Universal Robots URScript: FaiChun_9 Jan_2.script

def Machining2():
  # Default parameters:
  global speed_ms = 0.03
  global speed_rads = 0.75
  global accel_mss = 3
  global accel_radss = 1.2
  global blend_radius_m = 0.0003

  # Add subprograms here
  # Start of main program
  # Program generated by RoboDK v5.6.8 for UR10e on 09/01/2025 15:52:28
  # Using nominal kinematics.
  blend_radius_m = 0.0003
  speed_ms = 0.03
  # set_reference(p[0.335000, -0.075000, 0.000000, 0.000000, 0.000000, 0.000000])
  set_tcp(p[0.000000, 0.000000, 0.252000, 0.000000, 0.000000, 0.000000])
  # Show Tool
  movej([0.564339, -1.115693, -2.614907, -0.981789, 1.570796, 2.135135],accel_radss,speed_rads,0,blend_radius_m)
  movel([0.564339, -1.175740, -2.653333, -0.883316, 1.570796, 2.135135],accel_mss,speed_ms,0,blend_radius_m)
  #SetTool1
  #M_RunCode6
  #SetRPM60000
  speed_ms = 0.01
  #M_RunCode3
  movel([0.564339, -1.203294, -2.667921, -0.841174, 1.570796, 2.135135],accel_mss,speed_ms,0,blend_radius_m)
  speed_ms = 0.003
  movel([0.564339, -1.210543, -2.671504, -0.830343, 1.570796, 2.135135],accel_mss,speed_ms,0,blend_radius_m)
  speed_ms = 0.007
  movel([0.589071, -1.299862, -2.623221, -0.789306, 1.570796, 2.159867],accel_mss,speed_ms,0,blend_radius_m)
  movel([0.580877, -1.304600, -2.620384, -0.787405, 1.570796, 2.151673],accel_mss,speed_ms,0,blend_radius_m)
  movel([0.582153, -1.309303, -2.617539, -0.785547, 1.570796, 2.152950],accel_mss,speed_ms,0,blend_radius_m)
  movel([0.584262, -1.308090, -2.618275, -0.786023, 1.570796, 2.155058],accel_mss,speed_ms,0,blend_radius_m)
  movel([0.583431, -1.304986, -2.620151, -0.787251, 1.570796, 2.154228],accel_mss,speed_ms,0,blend_radius_m)
  movel([0.589492, -1.301500, -2.622244, -0.788646, 1.570796, 2.160288],accel_mss,speed_ms,0,blend_radius_m)
  movel([0.589686, -1.302254, -2.621792, -0.788342, 1.570796, 2.160482],accel_mss,speed_ms,0,blend_radius_m)
  movel([0.590691, -1.306131, -2.619461, -0.786797, 1.570796, 2.161487],accel_mss,speed_ms,0,blend_radius_m)
  movel([0.586616, -1.308460, -2.618051, -0.785878, 1.570796, 2.157412],accel_mss,speed_ms,0,blend_radius_m)
  movel([0.587040, -1.310068, -2.617073, -0.785248, 1.570796, 2.157837],accel_mss,speed_ms,0,blend_radius_m)
  movel([0.591108, -1.307752, -2.618481, -0.786157, 1.570796, 2.161905],accel_mss,speed_ms,0,blend_radius_m)
  movel([0.592288, -1.312350, -2.615680, -0.784359, 1.570796, 2.163085],accel_mss,speed_ms,0,blend_radius_m)
  movel([0.588242, -1.314642, -2.614274, -0.783473, 1.570796, 2.159038],accel_mss,speed_ms,0,blend_radius_m)
  movel([0.589043, -1.317715, -2.612378, -0.782297, 1.570796, 2.159840],accel_mss,speed_ms,0,blend_radius_m)
  movel([0.583100, -1.321078, -2.610288, -0.781023, 1.570796, 2.153897],accel_mss,speed_ms,0,blend_radius_m)
  movel([0.582276, -1.318031, -2.612181, -0.782176, 1.570796, 2.153073],accel_mss,speed_ms,0,blend_radius_m)
  movel([0.580193, -1.319220, -2.611444, -0.781725, 1.570796, 2.150989],accel_mss,speed_ms,0,blend_radius_m)
  movel([0.581023, -1.322259, -2.609550, -0.780580, 1.570796, 2.151819],accel_mss,speed_ms,0,blend_radius_m)
  movel([0.576077, -1.325076, -2.607784, -0.779529, 1.570796, 2.146874],accel_mss,speed_ms,0,blend_radius_m)
  movel([0.575122, -1.325624, -2.607439, -0.779326, 1.570796, 2.145918],accel_mss,speed_ms,0,blend_radius_m)
  movel([0.573856, -1.321163, -2.610235, -0.780991, 1.570796, 2.144653],accel_mss,speed_ms,0,blend_radius_m)
  movel([0.577859, -1.318861, -2.611667, -0.781861, 1.570796, 2.148656],accel_mss,speed_ms,0,blend_radius_m)
  movel([0.577420, -1.317283, -2.612645, -0.782461, 1.570796, 2.148217],accel_mss,speed_ms,0,blend_radius_m)
  movel([0.571335, -1.320792, -2.610466, -0.781131, 1.570796, 2.142131],accel_mss,speed_ms,0,blend_radius_m)
  movel([0.573058, -1.326803, -2.606696, -0.778890, 1.570796, 2.143854],accel_mss,speed_ms,0,blend_radius_m)
  movel([0.470799, -1.388192, -2.565343, -0.758854, 1.570796, 2.041595],accel_mss,speed_ms,0,blend_radius_m)
  movel([0.378716, -1.448552, -2.519372, -0.744466, 1.570796, 1.949513],accel_mss,speed_ms,0,blend_radius_m)
  movel([0.375919, -1.444184, -2.522882, -0.745323, 1.570796, 1.946716],accel_mss,speed_ms,0,blend_radius_m)
  movel([0.371026, -1.447561, -2.520170, -0.744657, 1.570796, 1.941822],accel_mss,speed_ms,0,blend_radius_m)
  movel([0.371758, -1.448686, -2.519263, -0.744440, 1.570796, 1.942554],accel_mss,speed_ms,0,blend_radius_m)
  movel([0.374972, -1.446470, -2.521049, -0.744871, 1.570796, 1.945769],accel_mss,speed_ms,0,blend_radius_m)
  movel([0.377041, -1.449694, -2.518449, -0.744246, 1.570796, 1.947837],accel_mss,speed_ms,0,blend_radius_m)
  movel([0.376268, -1.450223, -2.518020, -0.744145, 1.570796, 1.947064],accel_mss,speed_ms,0,blend_radius_m)
  movel([0.372297, -1.452950, -2.515807, -0.743632, 1.570796, 1.943093],accel_mss,speed_ms,0,blend_radius_m)
  movel([0.370895, -1.450790, -2.517562, -0.744037, 1.570796, 1.941691],accel_mss,speed_ms,0,blend_radius_m)
  movel([0.369236, -1.451936, -2.516632, -0.743821, 1.570796, 1.940032],accel_mss,speed_ms,0,blend_radius_m)
  movel([0.370642, -1.454090, -2.514879, -0.743420, 1.570796, 1.941438],accel_mss,speed_ms,0,blend_radius_m)
  movel([0.365939, -1.457337, -2.512222, -0.742829, 1.570796, 1.936735],accel_mss,speed_ms,0,blend_radius_m)
  movel([0.364521, -1.455203, -2.513970, -0.743216, 1.570796, 1.935317],accel_mss,speed_ms,0,blend_radius_m)
  movel([0.361355, -1.457405, -2.512167, -0.742817, 1.570796, 1.932152],accel_mss,speed_ms,0,blend_radius_m)
  movel([0.359234, -1.454259, -2.514741, -0.743389, 1.570796, 1.930031],accel_mss,speed_ms,0,blend_radius_m)
  movel([0.362410, -1.452037, -2.516550, -0.743802, 1.570796, 1.933206],accel_mss,speed_ms,0,blend_radius_m)
  movel([0.361665, -1.450927, -2.517450, -0.744011, 1.570796, 1.932462],accel_mss,speed_ms,0,blend_radius_m)
  movel([0.358487, -1.453153, -2.515642, -0.743594, 1.570796, 1.929284],accel_mss,speed_ms,0,blend_radius_m)
  movel([0.356688, -1.450515, -2.517784, -0.744090, 1.570796, 1.927484],accel_mss,speed_ms,0,blend_radius_m)
  movel([0.356339, -1.450002, -2.518199, -0.744187, 1.570796, 1.927136],accel_mss,speed_ms,0,blend_radius_m)
  movel([0.361066, -1.446678, -2.520881, -0.744830, 1.570796, 1.931863],accel_mss,speed_ms,0,blend_radius_m)
  movel([0.362508, -1.448824, -2.519152, -0.744413, 1.570796, 1.933304],accel_mss,speed_ms,0,blend_radius_m)
  movel([0.364168, -1.447664, -2.520088, -0.744637, 1.570796, 1.934964],accel_mss,speed_ms,0,blend_radius_m)
  movel([0.361980, -1.444391, -2.522716, -0.745282, 1.570796, 1.932777],accel_mss,speed_ms,0,blend_radius_m)
  movel([0.355583, -1.448897, -2.519093, -0.744399, 1.570796, 1.926379],accel_mss,speed_ms,0,blend_radius_m)
  movel([0.355230, -1.448386, -2.519506, -0.744497, 1.570796, 1.926027],accel_mss,speed_ms,0,blend_radius_m)
  movel([0.312755, -1.390773, -2.563487, -0.758128, 1.570796, 1.883551],accel_mss,speed_ms,0,blend_radius_m)
  movel([0.262445, -1.332364, -2.603164, -0.776861, 1.570796, 1.833241],accel_mss,speed_ms,0,blend_radius_m)
  movel([0.269473, -1.326239, -2.607051, -0.779098, 1.570796, 1.840270],accel_mss,speed_ms,0,blend_radius_m)
  movel([0.266416, -1.322928, -2.609132, -0.780329, 1.570796, 1.837212],accel_mss,speed_ms,0,blend_radius_m)
  movel([0.264580, -1.324533, -2.608125, -0.779731, 1.570796, 1.835377],accel_mss,speed_ms,0,blend_radius_m)
  movel([0.266599, -1.326703, -2.606759, -0.778927, 1.570796, 1.837395],accel_mss,speed_ms,0,blend_radius_m)
  movel([0.261398, -1.331241, -2.603881, -0.777267, 1.570796, 1.832194],accel_mss,speed_ms,0,blend_radius_m)
  movel([0.260914, -1.330724, -2.604210, -0.777455, 1.570796, 1.831710],accel_mss,speed_ms,0,blend_radius_m)
  movel([0.258394, -1.328064, -2.605899, -0.778426, 1.570796, 1.829190],accel_mss,speed_ms,0,blend_radius_m)
  movel([0.261907, -1.324978, -2.607845, -0.779565, 1.570796, 1.832703],accel_mss,speed_ms,0,blend_radius_m)
  movel([0.260849, -1.323857, -2.608550, -0.779982, 1.570796, 1.831646],accel_mss,speed_ms,0,blend_radius_m)
  movel([0.257334, -1.326952, -2.606602, -0.778835, 1.570796, 1.828131],accel_mss,speed_ms,0,blend_radius_m)
  movel([0.254293, -1.323782, -2.608597, -0.780010, 1.570796, 1.825090],accel_mss,speed_ms,0,blend_radius_m)
  movel([0.257815, -1.320661, -2.610547, -0.781180, 1.570796, 1.828612],accel_mss,speed_ms,0,blend_radius_m)
  movel([0.255752, -1.318503, -2.611889, -0.781997, 1.570796, 1.826548],accel_mss,speed_ms,0,blend_radius_m)
  movel([0.261012, -1.313833, -2.614771, -0.783785, 1.570796, 1.831808],accel_mss,speed_ms,0,blend_radius_m)
  movel([0.263069, -1.316016, -2.613428, -0.782946, 1.570796, 1.833865],accel_mss,speed_ms,0,blend_radius_m)
  movel([0.264921, -1.314382, -2.614434, -0.783573, 1.570796, 1.835718],accel_mss,speed_ms,0,blend_radius_m)
  movel([0.262867, -1.312190, -2.615778, -0.784421, 1.570796, 1.833663],accel_mss,speed_ms,0,blend_radius_m)
  movel([0.267321, -1.308250, -2.618179, -0.785961, 1.570796, 1.838117],accel_mss,speed_ms,0,blend_radius_m)
  movel([0.268189, -1.307485, -2.618642, -0.786262, 1.570796, 1.838985],accel_mss,speed_ms,0,blend_radius_m)
  movel([0.271218, -1.310771, -2.616645, -0.784973, 1.570796, 1.842014],accel_mss,speed_ms,0,blend_radius_m)
  movel([0.267627, -1.313924, -2.614715, -0.783750, 1.570796, 1.838423],accel_mss,speed_ms,0,blend_radius_m)
  movel([0.268684, -1.315067, -2.614012, -0.783310, 1.570796, 1.839480],accel_mss,speed_ms,0,blend_radius_m)
  movel([0.274144, -1.310287, -2.616940, -0.785162, 1.570796, 1.844940],accel_mss,speed_ms,0,blend_radius_m)
  movel([0.270069, -1.305826, -2.619645, -0.786918, 1.570796, 1.840865],accel_mss,speed_ms,0,blend_radius_m)
  movel([0.376357, -1.214643, -2.669493, -0.828252, 1.570796, 1.947154],accel_mss,speed_ms,0,blend_radius_m)
  movel([0.499980, -1.114188, -2.713609, -0.884591, 1.570796, 2.070776],accel_mss,speed_ms,0,blend_radius_m)
  movel([0.501179, -1.113243, -2.713976, -0.885169, 1.570796, 2.071975],accel_mss,speed_ms,0,blend_radius_m)
  movel([0.504077, -1.120540, -2.711120, -0.880729, 1.570796, 2.074873],accel_mss,speed_ms,0,blend_radius_m)
  movel([0.511634, -1.114642, -2.713433, -0.884314, 1.570796, 2.082430],accel_mss,speed_ms,0,blend_radius_m)
  movel([0.510904, -1.112724, -2.714178, -0.885487, 1.570796, 2.081700],accel_mss,speed_ms,0,blend_radius_m)
  movel([0.505914, -1.116627, -2.712658, -0.883104, 1.570796, 2.076710],accel_mss,speed_ms,0,blend_radius_m)
  movel([0.503784, -1.111195, -2.714769, -0.886425, 1.570796, 2.074581],accel_mss,speed_ms,0,blend_radius_m)
  movel([0.504986, -1.110247, -2.715135, -0.887007, 1.570796, 2.075782],accel_mss,speed_ms,0,blend_radius_m)
  movel([0.511228, -1.105329, -2.717019, -0.890042, 1.570796, 2.082024],accel_mss,speed_ms,0,blend_radius_m)
  movel([0.512639, -1.109056, -2.715593, -0.887740, 1.570796, 2.083436],accel_mss,speed_ms,0,blend_radius_m)
  movel([0.515254, -1.107012, -2.716376, -0.889001, 1.570796, 2.086050],accel_mss,speed_ms,0,blend_radius_m)
  movel([0.513852, -1.103266, -2.717802, -0.891321, 1.570796, 2.084649],accel_mss,speed_ms,0,blend_radius_m)
  movel([0.521382, -1.097360, -2.720023, -0.895006, 1.570796, 2.092179],accel_mss,speed_ms,0,blend_radius_m)
  movel([0.522759, -1.101158, -2.718598, -0.892633, 1.570796, 2.093556],accel_mss,speed_ms,0,blend_radius_m)
  movel([0.527861, -1.097189, -2.720087, -0.895113, 1.570796, 2.098658],accel_mss,speed_ms,0,blend_radius_m)
  movel([0.529846, -1.102848, -2.717960, -0.891581, 1.570796, 2.100643],accel_mss,speed_ms,0,blend_radius_m)
  movel([0.524769, -1.106765, -2.716471, -0.889153, 1.570796, 2.095565],accel_mss,speed_ms,0,blend_radius_m)
  movel([0.525468, -1.108724, -2.715721, -0.887945, 1.570796, 2.096264],accel_mss,speed_ms,0,blend_radius_m)
  movel([0.530535, -1.104825, -2.717210, -0.890354, 1.570796, 2.101331],accel_mss,speed_ms,0,blend_radius_m)
  movel([0.532478, -1.110454, -2.715055, -0.886880, 1.570796, 2.103274],accel_mss,speed_ms,0,blend_radius_m)
  movel([0.525035, -1.116137, -2.712849, -0.883402, 1.570796, 2.095831],accel_mss,speed_ms,0,blend_radius_m)
  movel([0.523692, -1.112395, -2.714305, -0.885689, 1.570796, 2.094489],accel_mss,speed_ms,0,blend_radius_m)
  movel([0.521088, -1.114399, -2.713527, -0.884462, 1.570796, 2.091884],accel_mss,speed_ms,0,blend_radius_m)
  movel([0.523134, -1.120056, -2.711311, -0.881022, 1.570796, 2.093931],accel_mss,speed_ms,0,blend_radius_m)
  movel([0.533154, -1.112420, -2.714296, -0.885673, 1.570796, 2.103950],accel_mss,speed_ms,0,blend_radius_m)
  movel([0.564339, -1.210543, -2.671504, -0.830343, 1.570796, 2.135135],accel_mss,speed_ms,0,blend_radius_m)
  speed_ms = 0.003
  movel([0.564339, -1.203294, -2.667921, -0.841174, 1.570796, 2.135135],accel_mss,speed_ms,0,blend_radius_m)
  speed_ms = 0.03
  movel([0.564339, -1.175740, -2.653333, -0.883316, 1.570796, 2.135135],accel_mss,speed_ms,0,blend_radius_m)
  #M_RunCode9
  movel([0.508673, -1.124915, -2.675707, -0.911767, 1.570796, 2.079469],accel_mss,speed_ms,0,blend_radius_m)
  #M_RunCode3
  movel([0.508673, -1.152779, -2.690963, -0.868647, 1.570796, 2.079469],accel_mss,speed_ms,0,blend_radius_m)
  speed_ms = 0.003
  movel([0.508673, -1.160141, -2.694716, -0.857531, 1.570796, 2.079469],accel_mss,speed_ms,0,blend_radius_m)
  speed_ms = 0.007
  movel([0.506502, -1.162157, -2.693839, -0.856392, 1.570796, 2.077298],accel_mss,speed_ms,0,blend_radius_m)
  movel([0.504257, -1.163601, -2.693209, -0.855579, 1.570796, 2.075054],accel_mss,speed_ms,0,blend_radius_m)
  movel([0.501934, -1.164482, -2.692823, -0.855084, 1.570796, 2.072730],accel_mss,speed_ms,0,blend_radius_m)
  movel([0.499527, -1.164799, -2.692684, -0.854906, 1.570796, 2.070323],accel_mss,speed_ms,0,blend_radius_m)
  movel([0.497561, -1.164580, -2.692780, -0.855029, 1.570796, 2.068358],accel_mss,speed_ms,0,blend_radius_m)
  movel([0.495980, -1.163844, -2.693102, -0.855442, 1.570796, 2.066776],accel_mss,speed_ms,0,blend_radius_m)
  movel([0.494731, -1.162733, -2.693588, -0.856068, 1.570796, 2.065527],accel_mss,speed_ms,0,blend_radius_m)
  movel([0.493766, -1.161377, -2.694179, -0.856833, 1.570796, 2.064563],accel_mss,speed_ms,0,blend_radius_m)
  movel([0.492038, -1.157449, -2.695881, -0.859059, 1.570796, 2.062834],accel_mss,speed_ms,0,blend_radius_m)
  movel([0.490361, -1.153755, -2.697467, -0.861167, 1.570796, 2.061158],accel_mss,speed_ms,0,blend_radius_m)
  movel([0.489477, -1.152506, -2.698000, -0.861883, 1.570796, 2.060274],accel_mss,speed_ms,0,blend_radius_m)
  movel([0.488348, -1.151492, -2.698432, -0.862465, 1.570796, 2.059144],accel_mss,speed_ms,0,blend_radius_m)
  movel([0.486938, -1.150837, -2.698710, -0.862842, 1.570796, 2.057734],accel_mss,speed_ms,0,blend_radius_m)
  movel([0.485211, -1.150668, -2.698782, -0.862939, 1.570796, 2.056007],accel_mss,speed_ms,0,blend_radius_m)
  movel([0.484699, -1.151781, -2.698309, -0.862299, 1.570796, 2.055495],accel_mss,speed_ms,0,blend_radius_m)
  movel([0.483417, -1.154849, -2.696999, -0.860541, 1.570796, 2.054213],accel_mss,speed_ms,0,blend_radius_m)
  movel([0.482581, -1.157515, -2.695853, -0.859021, 1.570796, 2.053377],accel_mss,speed_ms,0,blend_radius_m)
  movel([0.482187, -1.159786, -2.694871, -0.857732, 1.570796, 2.052983],accel_mss,speed_ms,0,blend_radius_m)
  movel([0.482229, -1.161669, -2.694052, -0.856668, 1.570796, 2.053026],accel_mss,speed_ms,0,blend_radius_m)
  movel([0.482647, -1.163187, -2.693390, -0.855812, 1.570796, 2.053443],accel_mss,speed_ms,0,blend_radius_m)
  movel([0.483386, -1.164368, -2.692873, -0.855148, 1.570796, 2.054183],accel_mss,speed_ms,0,blend_radius_m)
  movel([0.484448, -1.165208, -2.692505, -0.854677, 1.570796, 2.055244],accel_mss,speed_ms,0,blend_radius_m)
  movel([0.485828, -1.165715, -2.692281, -0.854392, 1.570796, 2.056624],accel_mss,speed_ms,0,blend_radius_m)
  movel([0.477331, -1.166016, -2.692149, -0.854224, 1.570796, 2.048127],accel_mss,speed_ms,0,blend_radius_m)
  movel([0.490968, -1.136326, -2.704766, -0.871297, 1.570796, 2.061764],accel_mss,speed_ms,0,blend_radius_m)
  movel([0.491843, -1.136290, -2.704781, -0.871318, 1.570796, 2.062639],accel_mss,speed_ms,0,blend_radius_m)
  movel([0.493898, -1.136547, -2.704675, -0.871167, 1.570796, 2.064694],accel_mss,speed_ms,0,blend_radius_m)
  movel([0.495585, -1.137510, -2.704280, -0.870600, 1.570796, 2.066381],accel_mss,speed_ms,0,blend_radius_m)
  movel([0.496938, -1.138969, -2.703678, -0.869741, 1.570796, 2.067734],accel_mss,speed_ms,0,blend_radius_m)
  movel([0.497990, -1.140717, -2.702955, -0.868716, 1.570796, 2.068786],accel_mss,speed_ms,0,blend_radius_m)
  movel([0.500129, -1.145961, -2.700769, -0.865660, 1.570796, 2.070926],accel_mss,speed_ms,0,blend_radius_m)
  movel([0.502024, -1.150859, -2.698701, -0.862829, 1.570796, 2.072821],accel_mss,speed_ms,0,blend_radius_m)
  movel([0.502966, -1.152496, -2.698005, -0.861888, 1.570796, 2.073762],accel_mss,speed_ms,0,blend_radius_m)
  movel([0.504145, -1.153842, -2.697430, -0.861117, 1.570796, 2.074941],accel_mss,speed_ms,0,blend_radius_m)
  movel([0.505585, -1.154734, -2.697048, -0.860607, 1.570796, 2.076381],accel_mss,speed_ms,0,blend_radius_m)
  movel([0.507301, -1.155017, -2.696927, -0.860445, 1.570796, 2.078097],accel_mss,speed_ms,0,blend_radius_m)
  movel([0.509687, -1.154592, -2.697109, -0.860688, 1.570796, 2.080483],accel_mss,speed_ms,0,blend_radius_m)
  movel([0.510798, -1.154086, -2.697325, -0.860977, 1.570796, 2.081594],accel_mss,speed_ms,0,blend_radius_m)
  movel([0.511860, -1.153380, -2.697627, -0.861382, 1.570796, 2.082656],accel_mss,speed_ms,0,blend_radius_m)
  movel([0.513679, -1.151630, -2.698373, -0.862386, 1.570796, 2.084475],accel_mss,speed_ms,0,blend_radius_m)
  movel([0.514984, -1.149603, -2.699233, -0.863553, 1.570796, 2.085781],accel_mss,speed_ms,0,blend_radius_m)
  movel([0.515524, -1.148232, -2.699813, -0.864344, 1.570796, 2.086320],accel_mss,speed_ms,0,blend_radius_m)
  movel([0.515638, -1.147219, -2.700240, -0.864930, 1.570796, 2.086434],accel_mss,speed_ms,0,blend_radius_m)
  movel([0.515378, -1.146593, -2.700503, -0.865293, 1.570796, 2.086174],accel_mss,speed_ms,0,blend_radius_m)
  movel([0.514794, -1.146390, -2.700588, -0.865411, 1.570796, 2.085591],accel_mss,speed_ms,0,blend_radius_m)
  movel([0.513538, -1.146896, -2.700375, -0.865117, 1.570796, 2.084335],accel_mss,speed_ms,0,blend_radius_m)
  movel([0.512295, -1.147497, -2.700123, -0.864769, 1.570796, 2.083092],accel_mss,speed_ms,0,blend_radius_m)
  movel([0.510910, -1.147730, -2.700025, -0.864635, 1.570796, 2.081706],accel_mss,speed_ms,0,blend_radius_m)
  movel([0.509562, -1.147401, -2.700163, -0.864825, 1.570796, 2.080359],accel_mss,speed_ms,0,blend_radius_m)
  movel([0.508936, -1.146367, -2.700598, -0.865424, 1.570796, 2.079732],accel_mss,speed_ms,0,blend_radius_m)
  movel([0.508971, -1.144842, -2.701238, -0.866310, 1.570796, 2.079767],accel_mss,speed_ms,0,blend_radius_m)
  movel([0.509601, -1.143041, -2.701990, -0.867358, 1.570796, 2.080397],accel_mss,speed_ms,0,blend_radius_m)
  movel([0.510703, -1.141227, -2.702744, -0.868418, 1.570796, 2.081499],accel_mss,speed_ms,0,blend_radius_m)
  movel([0.512151, -1.139669, -2.703389, -0.869331, 1.570796, 2.082947],accel_mss,speed_ms,0,blend_radius_m)
  movel([0.513800, -1.138587, -2.703836, -0.869966, 1.570796, 2.084597],accel_mss,speed_ms,0,blend_radius_m)
  movel([0.515498, -1.138213, -2.703990, -0.870186, 1.570796, 2.086294],accel_mss,speed_ms,0,blend_radius_m)
  movel([0.516742, -1.138401, -2.703913, -0.870075, 1.570796, 2.087539],accel_mss,speed_ms,0,blend_radius_m)
  movel([0.517622, -1.139001, -2.703665, -0.869722, 1.570796, 2.088419],accel_mss,speed_ms,0,blend_radius_m)
  movel([0.518134, -1.140018, -2.703245, -0.869126, 1.570796, 2.088931],accel_mss,speed_ms,0,blend_radius_m)
  movel([0.518284, -1.141439, -2.702656, -0.868294, 1.570796, 2.089081],accel_mss,speed_ms,0,blend_radius_m)
  movel([0.518110, -1.143170, -2.701936, -0.867283, 1.570796, 2.088906],accel_mss,speed_ms,0,blend_radius_m)
  movel([0.517640, -1.145109, -2.701126, -0.866154, 1.570796, 2.088437],accel_mss,speed_ms,0,blend_radius_m)
  movel([0.515835, -1.149598, -2.699236, -0.863556, 1.570796, 2.086632],accel_mss,speed_ms,0,blend_radius_m)
  movel([0.514301, -1.152485, -2.698009, -0.861894, 1.570796, 2.085098],accel_mss,speed_ms,0,blend_radius_m)
  movel([0.512598, -1.155205, -2.696846, -0.860338, 1.570796, 2.083394],accel_mss,speed_ms,0,blend_radius_m)
  movel([0.510722, -1.157753, -2.695750, -0.858886, 1.570796, 2.081518],accel_mss,speed_ms,0,blend_radius_m)
  movel([0.508673, -1.160141, -2.694716, -0.857531, 1.570796, 2.079469],accel_mss,speed_ms,0,blend_radius_m)
  speed_ms = 0.003
  movel([0.508673, -1.152779, -2.690963, -0.868647, 1.570796, 2.079469],accel_mss,speed_ms,0,blend_radius_m)
  speed_ms = 0.03
  movel([0.508673, -1.124915, -2.675707, -0.911767, 1.570796, 2.079469],accel_mss,speed_ms,0,blend_radius_m)
  #M_RunCode9
  movel([0.497081, -1.144256, -2.667496, -0.900636, 1.570796, 2.067877],accel_mss,speed_ms,0,blend_radius_m)
  #M_RunCode3
  movel([0.497081, -1.172027, -2.682500, -0.857862, 1.570796, 2.067877],accel_mss,speed_ms,0,blend_radius_m)
  speed_ms = 0.003
  movel([0.497081, -1.179353, -2.686188, -0.846848, 1.570796, 2.067877],accel_mss,speed_ms,0,blend_radius_m)
  speed_ms = 0.007
  movel([0.498395, -1.179888, -2.685945, -0.846556, 1.570796, 2.069191],accel_mss,speed_ms,0,blend_radius_m)
  movel([0.499154, -1.180637, -2.685604, -0.846148, 1.570796, 2.069950],accel_mss,speed_ms,0,blend_radius_m)
  movel([0.499362, -1.181606, -2.685163, -0.845621, 1.570796, 2.070158],accel_mss,speed_ms,0,blend_radius_m)
  movel([0.499017, -1.182788, -2.684622, -0.844979, 1.570796, 2.069813],accel_mss,speed_ms,0,blend_radius_m)
  movel([0.498226, -1.183973, -2.684079, -0.844337, 1.570796, 2.069022],accel_mss,speed_ms,0,blend_radius_m)
  movel([0.497089, -1.184946, -2.683632, -0.843811, 1.570796, 2.067885],accel_mss,speed_ms,0,blend_radius_m)
  movel([0.495612, -1.185707, -2.683282, -0.843400, 1.570796, 2.066408],accel_mss,speed_ms,0,blend_radius_m)
  movel([0.493784, -1.186265, -2.683025, -0.843099, 1.570796, 2.064581],accel_mss,speed_ms,0,blend_radius_m)
  movel([0.488939, -1.186979, -2.682695, -0.842715, 1.570796, 2.059736],accel_mss,speed_ms,0,blend_radius_m)
  movel([0.482396, -1.187317, -2.682539, -0.842533, 1.570796, 2.053192],accel_mss,speed_ms,0,blend_radius_m)
  movel([0.476031, -1.187267, -2.682562, -0.842560, 1.570796, 2.046827],accel_mss,speed_ms,0,blend_radius_m)
  movel([0.471758, -1.186758, -2.682797, -0.842834, 1.570796, 2.042555],accel_mss,speed_ms,0,blend_radius_m)
  movel([0.470420, -1.186270, -2.683022, -0.843096, 1.570796, 2.041216],accel_mss,speed_ms,0,blend_radius_m)
  movel([0.469629, -1.185561, -2.683349, -0.843479, 1.570796, 2.040426],accel_mss,speed_ms,0,blend_radius_m)
  movel([0.469386, -1.184621, -2.683782, -0.843986, 1.570796, 2.040183],accel_mss,speed_ms,0,blend_radius_m)
  movel([0.469698, -1.183447, -2.684320, -0.844621, 1.570796, 2.040494],accel_mss,speed_ms,0,blend_radius_m)
  movel([0.470461, -1.182257, -2.684865, -0.845267, 1.570796, 2.041257],accel_mss,speed_ms,0,blend_radius_m)
  movel([0.471587, -1.181260, -2.685321, -0.845809, 1.570796, 2.042384],accel_mss,speed_ms,0,blend_radius_m)
  movel([0.473070, -1.180460, -2.685685, -0.846244, 1.570796, 2.043867],accel_mss,speed_ms,0,blend_radius_m)
  movel([0.474917, -1.179854, -2.685960, -0.846575, 1.570796, 2.045714],accel_mss,speed_ms,0,blend_radius_m)
  movel([0.479828, -1.179041, -2.686329, -0.847018, 1.570796, 2.050624],accel_mss,speed_ms,0,blend_radius_m)
  movel([0.486445, -1.178651, -2.686507, -0.847232, 1.570796, 2.057241],accel_mss,speed_ms,0,blend_radius_m)
  movel([0.492832, -1.178747, -2.686463, -0.847179, 1.570796, 2.063629],accel_mss,speed_ms,0,blend_radius_m)
  movel([0.497081, -1.179353, -2.686188, -0.846848, 1.570796, 2.067877],accel_mss,speed_ms,0,blend_radius_m)
  speed_ms = 0.003
  movel([0.497081, -1.172027, -2.682500, -0.857862, 1.570796, 2.067877],accel_mss,speed_ms,0,blend_radius_m)
  speed_ms = 0.03
  movel([0.497081, -1.144256, -2.667496, -0.900636, 1.570796, 2.067877],accel_mss,speed_ms,0,blend_radius_m)
  #M_RunCode9
  movel([0.501396, -1.142283, -2.668351, -0.901755, 1.570796, 2.072192],accel_mss,speed_ms,0,blend_radius_m)
  #M_RunCode3
  movel([0.501396, -1.170065, -2.683380, -0.858944, 1.570796, 2.072192],accel_mss,speed_ms,0,blend_radius_m)
  speed_ms = 0.003
  movel([0.501396, -1.177394, -2.687075, -0.847919, 1.570796, 2.072192],accel_mss,speed_ms,0,blend_radius_m)
  speed_ms = 0.007
  movel([0.501126, -1.179098, -2.686304, -0.846987, 1.570796, 2.071922],accel_mss,speed_ms,0,blend_radius_m)
  movel([0.500589, -1.180897, -2.685486, -0.846006, 1.570796, 2.071385],accel_mss,speed_ms,0,blend_radius_m)
  movel([0.499790, -1.182783, -2.684624, -0.844981, 1.570796, 2.070587],accel_mss,speed_ms,0,blend_radius_m)
  movel([0.498777, -1.184668, -2.683760, -0.843961, 1.570796, 2.069573],accel_mss,speed_ms,0,blend_radius_m)
  movel([0.497593, -1.186454, -2.682938, -0.842998, 1.570796, 2.068389],accel_mss,speed_ms,0,blend_radius_m)
  movel([0.496241, -1.188138, -2.682158, -0.842092, 1.570796, 2.067037],accel_mss,speed_ms,0,blend_radius_m)
  movel([0.494719, -1.189727, -2.681421, -0.841241, 1.570796, 2.065515],accel_mss,speed_ms,0,blend_radius_m)
  movel([0.493045, -1.191188, -2.680740, -0.840460, 1.570796, 2.063841],accel_mss,speed_ms,0,blend_radius_m)
  movel([0.491239, -1.192488, -2.680133, -0.839768, 1.570796, 2.062036],accel_mss,speed_ms,0,blend_radius_m)
  movel([0.489295, -1.193633, -2.679596, -0.839160, 1.570796, 2.060092],accel_mss,speed_ms,0,blend_radius_m)
  movel([0.487213, -1.194624, -2.679131, -0.838635, 1.570796, 2.058010],accel_mss,speed_ms,0,blend_radius_m)
  movel([0.485034, -1.195426, -2.678753, -0.838210, 1.570796, 2.055830],accel_mss,speed_ms,0,blend_radius_m)
  movel([0.482787, -1.196014, -2.678476, -0.837899, 1.570796, 2.053583],accel_mss,speed_ms,0,blend_radius_m)
  movel([0.480475, -1.196388, -2.678299, -0.837702, 1.570796, 2.051271],accel_mss,speed_ms,0,blend_radius_m)
  movel([0.478097, -1.196547, -2.678224, -0.837618, 1.570796, 2.048893],accel_mss,speed_ms,0,blend_radius_m)
  movel([0.475817, -1.196490, -2.678251, -0.837648, 1.570796, 2.046613],accel_mss,speed_ms,0,blend_radius_m)
  movel([0.473808, -1.196212, -2.678382, -0.837795, 1.570796, 2.044604],accel_mss,speed_ms,0,blend_radius_m)
  movel([0.472068, -1.195712, -2.678618, -0.838059, 1.570796, 2.042864],accel_mss,speed_ms,0,blend_radius_m)
  movel([0.470598, -1.194990, -2.678958, -0.838441, 1.570796, 2.041394],accel_mss,speed_ms,0,blend_radius_m)
  movel([0.469404, -1.194073, -2.679390, -0.838926, 1.570796, 2.040200],accel_mss,speed_ms,0,blend_radius_m)
  movel([0.468492, -1.192991, -2.679897, -0.839500, 1.570796, 2.039288],accel_mss,speed_ms,0,blend_radius_m)
  movel([0.467863, -1.191747, -2.680479, -0.840162, 1.570796, 2.038659],accel_mss,speed_ms,0,blend_radius_m)
  movel([0.467519, -1.190332, -2.681140, -0.840918, 1.570796, 2.038316],accel_mss,speed_ms,0,blend_radius_m)
  movel([0.467450, -1.188781, -2.681861, -0.841747, 1.570796, 2.038247],accel_mss,speed_ms,0,blend_radius_m)
  movel([0.467649, -1.187124, -2.682628, -0.842637, 1.570796, 2.038445],accel_mss,speed_ms,0,blend_radius_m)
  movel([0.468121, -1.185356, -2.683444, -0.843589, 1.570796, 2.038917],accel_mss,speed_ms,0,blend_radius_m)
  movel([0.468861, -1.183480, -2.684305, -0.844604, 1.570796, 2.039658],accel_mss,speed_ms,0,blend_radius_m)
  movel([0.469829, -1.181592, -2.685169, -0.845628, 1.570796, 2.040626],accel_mss,speed_ms,0,blend_radius_m)
  movel([0.470983, -1.179781, -2.685994, -0.846614, 1.570796, 2.041779],accel_mss,speed_ms,0,blend_radius_m)
  movel([0.472326, -1.178055, -2.686777, -0.847558, 1.570796, 2.043122],accel_mss,speed_ms,0,blend_radius_m)
  movel([0.473857, -1.176411, -2.687519, -0.848459, 1.570796, 2.044653],accel_mss,speed_ms,0,blend_radius_m)
  movel([0.475556, -1.174883, -2.688207, -0.849299, 1.570796, 2.046352],accel_mss,speed_ms,0,blend_radius_m)
  movel([0.477400, -1.173508, -2.688824, -0.850058, 1.570796, 2.048196],accel_mss,speed_ms,0,blend_radius_m)
  movel([0.479390, -1.172291, -2.689368, -0.850730, 1.570796, 2.050187],accel_mss,speed_ms,0,blend_radius_m)
  movel([0.481526, -1.171228, -2.689842, -0.851319, 1.570796, 2.052322],accel_mss,speed_ms,0,blend_radius_m)
  movel([0.483771, -1.170360, -2.690228, -0.851801, 1.570796, 2.054567],accel_mss,speed_ms,0,blend_radius_m)
  movel([0.486082, -1.169720, -2.690512, -0.852157, 1.570796, 2.056878],accel_mss,speed_ms,0,blend_radius_m)
  movel([0.488460, -1.169311, -2.690694, -0.852384, 1.570796, 2.059257],accel_mss,speed_ms,0,blend_radius_m)
  movel([0.490905, -1.169136, -2.690771, -0.852481, 1.570796, 2.061701],accel_mss,speed_ms,0,blend_radius_m)
  movel([0.493234, -1.169201, -2.690742, -0.852445, 1.570796, 2.064030],accel_mss,speed_ms,0,blend_radius_m)
  movel([0.495277, -1.169508, -2.690606, -0.852275, 1.570796, 2.066073],accel_mss,speed_ms,0,blend_radius_m)
  movel([0.497033, -1.170056, -2.690363, -0.851970, 1.570796, 2.067829],accel_mss,speed_ms,0,blend_radius_m)
  movel([0.498501, -1.170839, -2.690015, -0.851535, 1.570796, 2.069297],accel_mss,speed_ms,0,blend_radius_m)
  movel([0.499675, -1.171826, -2.689575, -0.850988, 1.570796, 2.070472],accel_mss,speed_ms,0,blend_radius_m)
  movel([0.500550, -1.172979, -2.689060, -0.850350, 1.570796, 2.071346],accel_mss,speed_ms,0,blend_radius_m)
  movel([0.501123, -1.174299, -2.688469, -0.849621, 1.570796, 2.071919],accel_mss,speed_ms,0,blend_radius_m)
  movel([0.501400, -1.175784, -2.687802, -0.848804, 1.570796, 2.072196],accel_mss,speed_ms,0,blend_radius_m)
  movel([0.501396, -1.177394, -2.687075, -0.847919, 1.570796, 2.072192],accel_mss,speed_ms,0,blend_radius_m)
  speed_ms = 0.003
  movel([0.501396, -1.170065, -2.683380, -0.858944, 1.570796, 2.072192],accel_mss,speed_ms,0,blend_radius_m)
  speed_ms = 0.03
  movel([0.501396, -1.142283, -2.668351, -0.901755, 1.570796, 2.072192],accel_mss,speed_ms,0,blend_radius_m)
  #M_RunCode9
  movel([0.378486, -1.364194, -2.544953, -0.803242, 1.570796, 1.949283],accel_mss,speed_ms,0,blend_radius_m)
  #M_RunCode3
  movel([0.378486, -1.389086, -2.557074, -0.766230, 1.570796, 1.949283],accel_mss,speed_ms,0,blend_radius_m)
  speed_ms = 0.003
  movel([0.378486, -1.395545, -2.560031, -0.756813, 1.570796, 1.949283],accel_mss,speed_ms,0,blend_radius_m)
  speed_ms = 0.007
  movel([0.380119, -1.395727, -2.559899, -0.756763, 1.570796, 1.950915],accel_mss,speed_ms,0,blend_radius_m)
  movel([0.381530, -1.396365, -2.559434, -0.756590, 1.570796, 1.952326],accel_mss,speed_ms,0,blend_radius_m)
  movel([0.382726, -1.397324, -2.558734, -0.756330, 1.570796, 1.953523],accel_mss,speed_ms,0,blend_radius_m)
  movel([0.383717, -1.398472, -2.557895, -0.756022, 1.570796, 1.954513],accel_mss,speed_ms,0,blend_radius_m)
  movel([0.385894, -1.401918, -2.555364, -0.755107, 1.570796, 1.956690],accel_mss,speed_ms,0,blend_radius_m)
  movel([0.387854, -1.405140, -2.552982, -0.754268, 1.570796, 1.958650],accel_mss,speed_ms,0,blend_radius_m)
  movel([0.388748, -1.406222, -2.552178, -0.753989, 1.570796, 1.959544],accel_mss,speed_ms,0,blend_radius_m)
  movel([0.389806, -1.407111, -2.551517, -0.753761, 1.570796, 1.960602],accel_mss,speed_ms,0,blend_radius_m)
  movel([0.391022, -1.407700, -2.551078, -0.753611, 1.570796, 1.961819],accel_mss,speed_ms,0,blend_radius_m)
  movel([0.392399, -1.407890, -2.550936, -0.753563, 1.570796, 1.963195],accel_mss,speed_ms,0,blend_radius_m)
  movel([0.394233, -1.407617, -2.551140, -0.753632, 1.570796, 1.965029],accel_mss,speed_ms,0,blend_radius_m)
  movel([0.395059, -1.407284, -2.551388, -0.753717, 1.570796, 1.965855],accel_mss,speed_ms,0,blend_radius_m)
  movel([0.395827, -1.406821, -2.551733, -0.753836, 1.570796, 1.966623],accel_mss,speed_ms,0,blend_radius_m)
  movel([0.397082, -1.405675, -2.552584, -0.754129, 1.570796, 1.967879],accel_mss,speed_ms,0,blend_radius_m)
  movel([0.397912, -1.404346, -2.553570, -0.754473, 1.570796, 1.968708],accel_mss,speed_ms,0,blend_radius_m)
  movel([0.398201, -1.403448, -2.554234, -0.754706, 1.570796, 1.968997],accel_mss,speed_ms,0,blend_radius_m)
  movel([0.398192, -1.402782, -2.554726, -0.754880, 1.570796, 1.968988],accel_mss,speed_ms,0,blend_radius_m)
  movel([0.397925, -1.402374, -2.555028, -0.754987, 1.570796, 1.968721],accel_mss,speed_ms,0,blend_radius_m)
  movel([0.397445, -1.402238, -2.555128, -0.755023, 1.570796, 1.968242],accel_mss,speed_ms,0,blend_radius_m)
  movel([0.396511, -1.402568, -2.554885, -0.754937, 1.570796, 1.967307],accel_mss,speed_ms,0,blend_radius_m)
  movel([0.395591, -1.402959, -2.554596, -0.754834, 1.570796, 1.966388],accel_mss,speed_ms,0,blend_radius_m)
  movel([0.394526, -1.403109, -2.554485, -0.754795, 1.570796, 1.965322],accel_mss,speed_ms,0,blend_radius_m)
  movel([0.393436, -1.402891, -2.554646, -0.754852, 1.570796, 1.964232],accel_mss,speed_ms,0,blend_radius_m)
  movel([0.392846, -1.402211, -2.555148, -0.755030, 1.570796, 1.963642],accel_mss,speed_ms,0,blend_radius_m)
  movel([0.392723, -1.401214, -2.555882, -0.755293, 1.570796, 1.963520],accel_mss,speed_ms,0,blend_radius_m)
  movel([0.393041, -1.400035, -2.556749, -0.755605, 1.570796, 1.963837],accel_mss,speed_ms,0,blend_radius_m)
  movel([0.393730, -1.398853, -2.557616, -0.755920, 1.570796, 1.964527],accel_mss,speed_ms,0,blend_radius_m)
  movel([0.394713, -1.397839, -2.558358, -0.756192, 1.570796, 1.965509],accel_mss,speed_ms,0,blend_radius_m)
  movel([0.395898, -1.397138, -2.558870, -0.756381, 1.570796, 1.966694],accel_mss,speed_ms,0,blend_radius_m)
  movel([0.397191, -1.396897, -2.559046, -0.756446, 1.570796, 1.967988],accel_mss,speed_ms,0,blend_radius_m)
  movel([0.398186, -1.397023, -2.558954, -0.756412, 1.570796, 1.968982],accel_mss,speed_ms,0,blend_radius_m)
  movel([0.398934, -1.397418, -2.558666, -0.756305, 1.570796, 1.969730],accel_mss,speed_ms,0,blend_radius_m)
  movel([0.399440, -1.398079, -2.558182, -0.756127, 1.570796, 1.970236],accel_mss,speed_ms,0,blend_radius_m)
  movel([0.399697, -1.399009, -2.557502, -0.755878, 1.570796, 1.970494],accel_mss,speed_ms,0,blend_radius_m)
  movel([0.399730, -1.400139, -2.556673, -0.755577, 1.570796, 1.970526],accel_mss,speed_ms,0,blend_radius_m)
  movel([0.399553, -1.401406, -2.555741, -0.755242, 1.570796, 1.970349],accel_mss,speed_ms,0,blend_radius_m)
  movel([0.398578, -1.404344, -2.553572, -0.754473, 1.570796, 1.969374],accel_mss,speed_ms,0,blend_radius_m)
  movel([0.397658, -1.406238, -2.552166, -0.753985, 1.570796, 1.968454],accel_mss,speed_ms,0,blend_radius_m)
  movel([0.396583, -1.408023, -2.550837, -0.753529, 1.570796, 1.967380],accel_mss,speed_ms,0,blend_radius_m)
  movel([0.395357, -1.409701, -2.549583, -0.753105, 1.570796, 1.966154],accel_mss,speed_ms,0,blend_radius_m)
  movel([0.393975, -1.411273, -2.548405, -0.752712, 1.570796, 1.964771],accel_mss,speed_ms,0,blend_radius_m)
  movel([0.392460, -1.412604, -2.547403, -0.752381, 1.570796, 1.963256],accel_mss,speed_ms,0,blend_radius_m)
  movel([0.390831, -1.413556, -2.546686, -0.752147, 1.570796, 1.961627],accel_mss,speed_ms,0,blend_radius_m)
  movel([0.389086, -1.414133, -2.546251, -0.752005, 1.570796, 1.959883],accel_mss,speed_ms,0,blend_radius_m)
  movel([0.387222, -1.414339, -2.546095, -0.751955, 1.570796, 1.958019],accel_mss,speed_ms,0,blend_radius_m)
  movel([0.385652, -1.414186, -2.546210, -0.751992, 1.570796, 1.956448],accel_mss,speed_ms,0,blend_radius_m)
  movel([0.384339, -1.413696, -2.546581, -0.752112, 1.570796, 1.955135],accel_mss,speed_ms,0,blend_radius_m)
  movel([0.383252, -1.412953, -2.547141, -0.752295, 1.570796, 1.954048],accel_mss,speed_ms,0,blend_radius_m)
  movel([0.382365, -1.412051, -2.547819, -0.752518, 1.570796, 1.953161],accel_mss,speed_ms,0,blend_radius_m)
  movel([0.380633, -1.409448, -2.549772, -0.753169, 1.570796, 1.951429],accel_mss,speed_ms,0,blend_radius_m)
  movel([0.378972, -1.407001, -2.551598, -0.753789, 1.570796, 1.949768],accel_mss,speed_ms,0,blend_radius_m)
  movel([0.378159, -1.406171, -2.552216, -0.754002, 1.570796, 1.948956],accel_mss,speed_ms,0,blend_radius_m)
  movel([0.377180, -1.405497, -2.552717, -0.754175, 1.570796, 1.947977],accel_mss,speed_ms,0,blend_radius_m)
  movel([0.376010, -1.405059, -2.553041, -0.754288, 1.570796, 1.946807],accel_mss,speed_ms,0,blend_radius_m)
  movel([0.374641, -1.404938, -2.553131, -0.754320, 1.570796, 1.945437],accel_mss,speed_ms,0,blend_radius_m)
  movel([0.374343, -1.405668, -2.552589, -0.754131, 1.570796, 1.945139],accel_mss,speed_ms,0,blend_radius_m)
  movel([0.373624, -1.407683, -2.551090, -0.753616, 1.570796, 1.944421],accel_mss,speed_ms,0,blend_radius_m)
  movel([0.373215, -1.409441, -2.549777, -0.753170, 1.570796, 1.944011],accel_mss,speed_ms,0,blend_radius_m)
  movel([0.373114, -1.410945, -2.548651, -0.752794, 1.570796, 1.943910],accel_mss,speed_ms,0,blend_radius_m)
  movel([0.373319, -1.412193, -2.547713, -0.752483, 1.570796, 1.944115],accel_mss,speed_ms,0,blend_radius_m)
  movel([0.373789, -1.413203, -2.546952, -0.752234, 1.570796, 1.944585],accel_mss,speed_ms,0,blend_radius_m)
  movel([0.374478, -1.413989, -2.546360, -0.752040, 1.570796, 1.945275],accel_mss,speed_ms,0,blend_radius_m)
  movel([0.375390, -1.414554, -2.545933, -0.751902, 1.570796, 1.946186],accel_mss,speed_ms,0,blend_radius_m)
  movel([0.376523, -1.414896, -2.545674, -0.751819, 1.570796, 1.947320],accel_mss,speed_ms,0,blend_radius_m)
  movel([0.369870, -1.415050, -2.545557, -0.751781, 1.570796, 1.940666],accel_mss,speed_ms,0,blend_radius_m)
  movel([0.377808, -1.395563, -2.560018, -0.756808, 1.570796, 1.948604],accel_mss,speed_ms,0,blend_radius_m)
  movel([0.378486, -1.395545, -2.560031, -0.756813, 1.570796, 1.949283],accel_mss,speed_ms,0,blend_radius_m)
  speed_ms = 0.003
  movel([0.378486, -1.389086, -2.557074, -0.766230, 1.570796, 1.949283],accel_mss,speed_ms,0,blend_radius_m)
  speed_ms = 0.03
  movel([0.378486, -1.364194, -2.544953, -0.803242, 1.570796, 1.949283],accel_mss,speed_ms,0,blend_radius_m)
  #M_RunCode9
  movel([0.373054, -1.386537, -2.529095, -0.796757, 1.570796, 1.943850],accel_mss,speed_ms,0,blend_radius_m)
  #M_RunCode3
  movel([0.373054, -1.411000, -2.540935, -0.760454, 1.570796, 1.943850],accel_mss,speed_ms,0,blend_radius_m)
  speed_ms = 0.003
  movel([0.373054, -1.417339, -2.543822, -0.751228, 1.570796, 1.943850],accel_mss,speed_ms,0,blend_radius_m)
  speed_ms = 0.007
  movel([0.374143, -1.417539, -2.543670, -0.751180, 1.570796, 1.944939],accel_mss,speed_ms,0,blend_radius_m)
  movel([0.374760, -1.418189, -2.543176, -0.751024, 1.570796, 1.945557],accel_mss,speed_ms,0,blend_radius_m)
  movel([0.374917, -1.419156, -2.542439, -0.750794, 1.570796, 1.945713],accel_mss,speed_ms,0,blend_radius_m)
  movel([0.374633, -1.420296, -2.541569, -0.750524, 1.570796, 1.945429],accel_mss,speed_ms,0,blend_radius_m)
  movel([0.373980, -1.421442, -2.540692, -0.750255, 1.570796, 1.944776],accel_mss,speed_ms,0,blend_radius_m)
  movel([0.373026, -1.422424, -2.539939, -0.750026, 1.570796, 1.943823],accel_mss,speed_ms,0,blend_radius_m)
  movel([0.371867, -1.423108, -2.539413, -0.749867, 1.570796, 1.942663],accel_mss,speed_ms,0,blend_radius_m)
  movel([0.370603, -1.423355, -2.539224, -0.749810, 1.570796, 1.941400],accel_mss,speed_ms,0,blend_radius_m)
  movel([0.369670, -1.423239, -2.539313, -0.749837, 1.570796, 1.940466],accel_mss,speed_ms,0,blend_radius_m)
  movel([0.369080, -1.422882, -2.539587, -0.749920, 1.570796, 1.939877],accel_mss,speed_ms,0,blend_radius_m)
  movel([0.368422, -1.422586, -2.539815, -0.749988, 1.570796, 1.939218],accel_mss,speed_ms,0,blend_radius_m)
  movel([0.367836, -1.422738, -2.539698, -0.749953, 1.570796, 1.938632],accel_mss,speed_ms,0,blend_radius_m)
  movel([0.367230, -1.423163, -2.539371, -0.749854, 1.570796, 1.938026],accel_mss,speed_ms,0,blend_radius_m)
  movel([0.366694, -1.423770, -2.538905, -0.749714, 1.570796, 1.937491],accel_mss,speed_ms,0,blend_radius_m)
  movel([0.366316, -1.424471, -2.538365, -0.749553, 1.570796, 1.937112],accel_mss,speed_ms,0,blend_radius_m)
  movel([0.366043, -1.425391, -2.537656, -0.749343, 1.570796, 1.936839],accel_mss,speed_ms,0,blend_radius_m)
  movel([0.366002, -1.426224, -2.537012, -0.749153, 1.570796, 1.936799],accel_mss,speed_ms,0,blend_radius_m)
  movel([0.366192, -1.426968, -2.536436, -0.748985, 1.570796, 1.936989],accel_mss,speed_ms,0,blend_radius_m)
  movel([0.366611, -1.427630, -2.535924, -0.748836, 1.570796, 1.937407],accel_mss,speed_ms,0,blend_radius_m)
  movel([0.367235, -1.428165, -2.535509, -0.748716, 1.570796, 1.938032],accel_mss,speed_ms,0,blend_radius_m)
  movel([0.368038, -1.428539, -2.535218, -0.748632, 1.570796, 1.938834],accel_mss,speed_ms,0,blend_radius_m)
  movel([0.369018, -1.428754, -2.535051, -0.748584, 1.570796, 1.939814],accel_mss,speed_ms,0,blend_radius_m)
  movel([0.370176, -1.428809, -2.535008, -0.748572, 1.570796, 1.940973],accel_mss,speed_ms,0,blend_radius_m)
  movel([0.372277, -1.428488, -2.535257, -0.748643, 1.570796, 1.943073],accel_mss,speed_ms,0,blend_radius_m)
  movel([0.374406, -1.427607, -2.535941, -0.748841, 1.570796, 1.945202],accel_mss,speed_ms,0,blend_radius_m)
  movel([0.375468, -1.426949, -2.536451, -0.748989, 1.570796, 1.946265],accel_mss,speed_ms,0,blend_radius_m)
  movel([0.376504, -1.426147, -2.537071, -0.749171, 1.570796, 1.947300],accel_mss,speed_ms,0,blend_radius_m)
  movel([0.378505, -1.424090, -2.538658, -0.749641, 1.570796, 1.949302],accel_mss,speed_ms,0,blend_radius_m)
  movel([0.380333, -1.421463, -2.540676, -0.750250, 1.570796, 1.951130],accel_mss,speed_ms,0,blend_radius_m)
  movel([0.381903, -1.418285, -2.543103, -0.751001, 1.570796, 1.952700],accel_mss,speed_ms,0,blend_radius_m)
  movel([0.391997, -1.418198, -2.543169, -0.751022, 1.570796, 1.962793],accel_mss,speed_ms,0,blend_radius_m)
  movel([0.385959, -1.432381, -2.532223, -0.747785, 1.570796, 1.956755],accel_mss,speed_ms,0,blend_radius_m)
  movel([0.379469, -1.432425, -2.532188, -0.747775, 1.570796, 1.950266],accel_mss,speed_ms,0,blend_radius_m)
  movel([0.381244, -1.431876, -2.532618, -0.747895, 1.570796, 1.952041],accel_mss,speed_ms,0,blend_radius_m)
  movel([0.383068, -1.430883, -2.533394, -0.748113, 1.570796, 1.953864],accel_mss,speed_ms,0,blend_radius_m)
  movel([0.384851, -1.429490, -2.534478, -0.748420, 1.570796, 1.955647],accel_mss,speed_ms,0,blend_radius_m)
  movel([0.386501, -1.427748, -2.535832, -0.748809, 1.570796, 1.957298],accel_mss,speed_ms,0,blend_radius_m)
  movel([0.387947, -1.425706, -2.537412, -0.749271, 1.570796, 1.958743],accel_mss,speed_ms,0,blend_radius_m)
  movel([0.389111, -1.423424, -2.539171, -0.749794, 1.570796, 1.959907],accel_mss,speed_ms,0,blend_radius_m)
  movel([0.381698, -1.423483, -2.539126, -0.749781, 1.570796, 1.952494],accel_mss,speed_ms,0,blend_radius_m)
  movel([0.380319, -1.426295, -2.536957, -0.749137, 1.570796, 1.951116],accel_mss,speed_ms,0,blend_radius_m)
  movel([0.378590, -1.428985, -2.534872, -0.748533, 1.570796, 1.949387],accel_mss,speed_ms,0,blend_radius_m)
  movel([0.376562, -1.431371, -2.533012, -0.748006, 1.570796, 1.947358],accel_mss,speed_ms,0,blend_radius_m)
  movel([0.375453, -1.432385, -2.532219, -0.747784, 1.570796, 1.946249],accel_mss,speed_ms,0,blend_radius_m)
  movel([0.374283, -1.433281, -2.531518, -0.747590, 1.570796, 1.945080],accel_mss,speed_ms,0,blend_radius_m)
  movel([0.373065, -1.434017, -2.530941, -0.747431, 1.570796, 1.943862],accel_mss,speed_ms,0,blend_radius_m)
  movel([0.371820, -1.434547, -2.530524, -0.747317, 1.570796, 1.942616],accel_mss,speed_ms,0,blend_radius_m)
  movel([0.370542, -1.434876, -2.530266, -0.747247, 1.570796, 1.941339],accel_mss,speed_ms,0,blend_radius_m)
  movel([0.369238, -1.435001, -2.530168, -0.747220, 1.570796, 1.940034],accel_mss,speed_ms,0,blend_radius_m)
  movel([0.368011, -1.434929, -2.530224, -0.747236, 1.570796, 1.938807],accel_mss,speed_ms,0,blend_radius_m)
  movel([0.366967, -1.434666, -2.530431, -0.747292, 1.570796, 1.937764],accel_mss,speed_ms,0,blend_radius_m)
  movel([0.366110, -1.434210, -2.530789, -0.747390, 1.570796, 1.936907],accel_mss,speed_ms,0,blend_radius_m)
  movel([0.365439, -1.433562, -2.531298, -0.747529, 1.570796, 1.936235],accel_mss,speed_ms,0,blend_radius_m)
  movel([0.364597, -1.431859, -2.532631, -0.747899, 1.570796, 1.935394],accel_mss,speed_ms,0,blend_radius_m)
  movel([0.364385, -1.429734, -2.534289, -0.748366, 1.570796, 1.935181],accel_mss,speed_ms,0,blend_radius_m)
  movel([0.364715, -1.427351, -2.536140, -0.748898, 1.570796, 1.935512],accel_mss,speed_ms,0,blend_radius_m)
  movel([0.365497, -1.424883, -2.538048, -0.749459, 1.570796, 1.936293],accel_mss,speed_ms,0,blend_radius_m)
  movel([0.366314, -1.423176, -2.539361, -0.749851, 1.570796, 1.937110],accel_mss,speed_ms,0,blend_radius_m)
  movel([0.367412, -1.421439, -2.540694, -0.750256, 1.570796, 1.938209],accel_mss,speed_ms,0,blend_radius_m)
  movel([0.368714, -1.419835, -2.541921, -0.750633, 1.570796, 1.939510],accel_mss,speed_ms,0,blend_radius_m)
  movel([0.370145, -1.418530, -2.542916, -0.750943, 1.570796, 1.940941],accel_mss,speed_ms,0,blend_radius_m)
  movel([0.371620, -1.417653, -2.543584, -0.751152, 1.570796, 1.942416],accel_mss,speed_ms,0,blend_radius_m)
  movel([0.373054, -1.417339, -2.543822, -0.751228, 1.570796, 1.943850],accel_mss,speed_ms,0,blend_radius_m)
  speed_ms = 0.003
  movel([0.373054, -1.411000, -2.540935, -0.760454, 1.570796, 1.943850],accel_mss,speed_ms,0,blend_radius_m)
  speed_ms = 0.03
  movel([0.373054, -1.386537, -2.529095, -0.796757, 1.570796, 1.943850],accel_mss,speed_ms,0,blend_radius_m)
  #M_RunCode9
  movel([0.456957, -1.302684, -2.585134, -0.824571, 1.570796, 2.027753],accel_mss,speed_ms,0,blend_radius_m)
  #M_RunCode3
  movel([0.456957, -1.328657, -2.598047, -0.785686, 1.570796, 2.027753],accel_mss,speed_ms,0,blend_radius_m)
  speed_ms = 0.003
  movel([0.456957, -1.335424, -2.601204, -0.775762, 1.570796, 2.027753],accel_mss,speed_ms,0,blend_radius_m)
  speed_ms = 0.007
  movel([0.457043, -1.335364, -2.601242, -0.775783, 1.570796, 2.027839],accel_mss,speed_ms,0,blend_radius_m)
  movel([0.456957, -1.335424, -2.601204, -0.775762, 1.570796, 2.027753],accel_mss,speed_ms,0,blend_radius_m)
  speed_ms = 0.003
  movel([0.456957, -1.328657, -2.598047, -0.785686, 1.570796, 2.027753],accel_mss,speed_ms,0,blend_radius_m)
  speed_ms = 0.03
  movel([0.456957, -1.302684, -2.585134, -0.824571, 1.570796, 2.027753],accel_mss,speed_ms,0,blend_radius_m)
  #M_RunCode9
  movel([0.434206, -1.314146, -2.578022, -0.820220, 1.570796, 2.005002],accel_mss,speed_ms,0,blend_radius_m)
  #M_RunCode3
  movel([0.434206, -1.339930, -2.590785, -0.781673, 1.570796, 2.005002],accel_mss,speed_ms,0,blend_radius_m)
  speed_ms = 0.003
  movel([0.434206, -1.346643, -2.593905, -0.771842, 1.570796, 2.005002],accel_mss,speed_ms,0,blend_radius_m)
  speed_ms = 0.007
  movel([0.434230, -1.347825, -2.593125, -0.771438, 1.570796, 2.005027],accel_mss,speed_ms,0,blend_radius_m)
  movel([0.433916, -1.349258, -2.592178, -0.770953, 1.570796, 2.004712],accel_mss,speed_ms,0,blend_radius_m)
  movel([0.432901, -1.351412, -2.590749, -0.770228, 1.570796, 2.003697],accel_mss,speed_ms,0,blend_radius_m)
  movel([0.431373, -1.353297, -2.589494, -0.769598, 1.570796, 2.002170],accel_mss,speed_ms,0,blend_radius_m)
  movel([0.429428, -1.354894, -2.588426, -0.769069, 1.570796, 2.000224],accel_mss,speed_ms,0,blend_radius_m)
  movel([0.427164, -1.356179, -2.587564, -0.768646, 1.570796, 1.997960],accel_mss,speed_ms,0,blend_radius_m)
  movel([0.424569, -1.357112, -2.586937, -0.768340, 1.570796, 1.995365],accel_mss,speed_ms,0,blend_radius_m)
  movel([0.422436, -1.357318, -2.586798, -0.768273, 1.570796, 1.993232],accel_mss,speed_ms,0,blend_radius_m)
  movel([0.420729, -1.356905, -2.587076, -0.768408, 1.570796, 1.991525],accel_mss,speed_ms,0,blend_radius_m)
  movel([0.419414, -1.355971, -2.587704, -0.768714, 1.570796, 1.990210],accel_mss,speed_ms,0,blend_radius_m)
  movel([0.418455, -1.354624, -2.588607, -0.769158, 1.570796, 1.989252],accel_mss,speed_ms,0,blend_radius_m)
  movel([0.417823, -1.352963, -2.589717, -0.769710, 1.570796, 1.988619],accel_mss,speed_ms,0,blend_radius_m)
  movel([0.417486, -1.351092, -2.590962, -0.770335, 1.570796, 1.988282],accel_mss,speed_ms,0,blend_radius_m)
  movel([0.417413, -1.349115, -2.592273, -0.771001, 1.570796, 1.988210],accel_mss,speed_ms,0,blend_radius_m)
  movel([0.419866, -1.347321, -2.593458, -0.771610, 1.570796, 1.990662],accel_mss,speed_ms,0,blend_radius_m)
  movel([0.422769, -1.345812, -2.594451, -0.772126, 1.570796, 1.993565],accel_mss,speed_ms,0,blend_radius_m)
  movel([0.425843, -1.344709, -2.595175, -0.772505, 1.570796, 1.996640],accel_mss,speed_ms,0,blend_radius_m)
  movel([0.428805, -1.344126, -2.595557, -0.772706, 1.570796, 1.999601],accel_mss,speed_ms,0,blend_radius_m)
  movel([0.431375, -1.344181, -2.595521, -0.772687, 1.570796, 2.002171],accel_mss,speed_ms,0,blend_radius_m)
  movel([0.432423, -1.344484, -2.595323, -0.772583, 1.570796, 2.003219],accel_mss,speed_ms,0,blend_radius_m)
  movel([0.433268, -1.344985, -2.594994, -0.772410, 1.570796, 2.004064],accel_mss,speed_ms,0,blend_radius_m)
  movel([0.433873, -1.345700, -2.594524, -0.772164, 1.570796, 2.004669],accel_mss,speed_ms,0,blend_radius_m)
  movel([0.434206, -1.346643, -2.593905, -0.771842, 1.570796, 2.005002],accel_mss,speed_ms,0,blend_radius_m)
  speed_ms = 0.003
  movel([0.434206, -1.339930, -2.590785, -0.781673, 1.570796, 2.005002],accel_mss,speed_ms,0,blend_radius_m)
  speed_ms = 0.03
  movel([0.434206, -1.314146, -2.578022, -0.820220, 1.570796, 2.005002],accel_mss,speed_ms,0,blend_radius_m)
  #M_RunCode9
  movel([0.495621, -1.297461, -2.588320, -0.826609, 1.570796, 2.066418],accel_mss,speed_ms,0,blend_radius_m)
  #M_RunCode3
  movel([0.495621, -1.323517, -2.601300, -0.787571, 1.570796, 2.066418],accel_mss,speed_ms,0,blend_radius_m)
  speed_ms = 0.003
  movel([0.495621, -1.330309, -2.604474, -0.777606, 1.570796, 2.066418],accel_mss,speed_ms,0,blend_radius_m)
  speed_ms = 0.007
  movel([0.496230, -1.328877, -2.605383, -0.778128, 1.570796, 2.067026],accel_mss,speed_ms,0,blend_radius_m)
  movel([0.497032, -1.327417, -2.606308, -0.778664, 1.570796, 2.067828],accel_mss,speed_ms,0,blend_radius_m)
  movel([0.497406, -1.327643, -2.606165, -0.778581, 1.570796, 2.068202],accel_mss,speed_ms,0,blend_radius_m)
  movel([0.497374, -1.328119, -2.605864, -0.778406, 1.570796, 2.068170],accel_mss,speed_ms,0,blend_radius_m)
  movel([0.497378, -1.328653, -2.605526, -0.778211, 1.570796, 2.068174],accel_mss,speed_ms,0,blend_radius_m)
  movel([0.497857, -1.329054, -2.605271, -0.778064, 1.570796, 2.068654],accel_mss,speed_ms,0,blend_radius_m)
  movel([0.498655, -1.329140, -2.605217, -0.778032, 1.570796, 2.069452],accel_mss,speed_ms,0,blend_radius_m)
  movel([0.499556, -1.329032, -2.605285, -0.778072, 1.570796, 2.070353],accel_mss,speed_ms,0,blend_radius_m)
  movel([0.500825, -1.328832, -2.605412, -0.778145, 1.570796, 2.071622],accel_mss,speed_ms,0,blend_radius_m)
  movel([0.501916, -1.327012, -2.606564, -0.778813, 1.570796, 2.072712],accel_mss,speed_ms,0,blend_radius_m)
  movel([0.502401, -1.325471, -2.607535, -0.779383, 1.570796, 2.073197],accel_mss,speed_ms,0,blend_radius_m)
  movel([0.502337, -1.324859, -2.607920, -0.779610, 1.570796, 2.073133],accel_mss,speed_ms,0,blend_radius_m)
  movel([0.502031, -1.324383, -2.608220, -0.779787, 1.570796, 2.072828],accel_mss,speed_ms,0,blend_radius_m)
  movel([0.501449, -1.324062, -2.608421, -0.779906, 1.570796, 2.072245],accel_mss,speed_ms,0,blend_radius_m)
  movel([0.500560, -1.323923, -2.608508, -0.779958, 1.570796, 2.071356],accel_mss,speed_ms,0,blend_radius_m)
  movel([0.501570, -1.323058, -2.609051, -0.780281, 1.570796, 2.072366],accel_mss,speed_ms,0,blend_radius_m)
  movel([0.502493, -1.322400, -2.609462, -0.780527, 1.570796, 2.073290],accel_mss,speed_ms,0,blend_radius_m)
  movel([0.502874, -1.322255, -2.609553, -0.780581, 1.570796, 2.073670],accel_mss,speed_ms,0,blend_radius_m)
  movel([0.503173, -1.322286, -2.609534, -0.780570, 1.570796, 2.073970],accel_mss,speed_ms,0,blend_radius_m)
  movel([0.503455, -1.323044, -2.609059, -0.780286, 1.570796, 2.074252],accel_mss,speed_ms,0,blend_radius_m)
  movel([0.503269, -1.325026, -2.607815, -0.779548, 1.570796, 2.074065],accel_mss,speed_ms,0,blend_radius_m)
  movel([0.502577, -1.327171, -2.606464, -0.778755, 1.570796, 2.073374],accel_mss,speed_ms,0,blend_radius_m)
  movel([0.502021, -1.328201, -2.605812, -0.778376, 1.570796, 2.072817],accel_mss,speed_ms,0,blend_radius_m)
  movel([0.501308, -1.329152, -2.605209, -0.778028, 1.570796, 2.072104],accel_mss,speed_ms,0,blend_radius_m)
  movel([0.500430, -1.329980, -2.604683, -0.777726, 1.570796, 2.071227],accel_mss,speed_ms,0,blend_radius_m)
  movel([0.499378, -1.330648, -2.604259, -0.777483, 1.570796, 2.070174],accel_mss,speed_ms,0,blend_radius_m)
  movel([0.499440, -1.329425, -2.605036, -0.777928, 1.570796, 2.070236],accel_mss,speed_ms,0,blend_radius_m)
  movel([0.495661, -1.332838, -2.602861, -0.776690, 1.570796, 2.066457],accel_mss,speed_ms,0,blend_radius_m)
  movel([0.495376, -1.331650, -2.603620, -0.777119, 1.570796, 2.066172],accel_mss,speed_ms,0,blend_radius_m)
  movel([0.495621, -1.330309, -2.604474, -0.777606, 1.570796, 2.066418],accel_mss,speed_ms,0,blend_radius_m)
  speed_ms = 0.003
  movel([0.495621, -1.323517, -2.601300, -0.787571, 1.570796, 2.066418],accel_mss,speed_ms,0,blend_radius_m)
  speed_ms = 0.03
  movel([0.495621, -1.297461, -2.588320, -0.826609, 1.570796, 2.066418],accel_mss,speed_ms,0,blend_radius_m)
  #M_RunCode9
  movel([0.511194, -1.258845, -2.610818, -0.842726, 1.570796, 2.081990],accel_mss,speed_ms,0,blend_radius_m)
  #M_RunCode3
  movel([0.511194, -1.285477, -2.624306, -0.802605, 1.570796, 2.081990],accel_mss,speed_ms,0,blend_radius_m)
  speed_ms = 0.003
  movel([0.511194, -1.292438, -2.627609, -0.792342, 1.570796, 2.081990],accel_mss,speed_ms,0,blend_radius_m)
  speed_ms = 0.007
  movel([0.509391, -1.292526, -2.627557, -0.792306, 1.570796, 2.080187],accel_mss,speed_ms,0,blend_radius_m)
  movel([0.507674, -1.292384, -2.627640, -0.792365, 1.570796, 2.078471],accel_mss,speed_ms,0,blend_radius_m)
  movel([0.506070, -1.292003, -2.627863, -0.792522, 1.570796, 2.076867],accel_mss,speed_ms,0,blend_radius_m)
  movel([0.504607, -1.291371, -2.628233, -0.792784, 1.570796, 2.075403],accel_mss,speed_ms,0,blend_radius_m)
  movel([0.503311, -1.290484, -2.628752, -0.793154, 1.570796, 2.074107],accel_mss,speed_ms,0,blend_radius_m)
  movel([0.502827, -1.289811, -2.629144, -0.793434, 1.570796, 2.073623],accel_mss,speed_ms,0,blend_radius_m)
  movel([0.502472, -1.288966, -2.629636, -0.793787, 1.570796, 2.073269],accel_mss,speed_ms,0,blend_radius_m)
  movel([0.502151, -1.288211, -2.630075, -0.794103, 1.570796, 2.072948],accel_mss,speed_ms,0,blend_radius_m)
  movel([0.501756, -1.287808, -2.630309, -0.794272, 1.570796, 2.072553],accel_mss,speed_ms,0,blend_radius_m)
  movel([0.500573, -1.287809, -2.630309, -0.794272, 1.570796, 2.071369],accel_mss,speed_ms,0,blend_radius_m)
  movel([0.498809, -1.288086, -2.630147, -0.794155, 1.570796, 2.069605],accel_mss,speed_ms,0,blend_radius_m)
  movel([0.496952, -1.288406, -2.629962, -0.794021, 1.570796, 2.067748],accel_mss,speed_ms,0,blend_radius_m)
  movel([0.495490, -1.288524, -2.629893, -0.793972, 1.570796, 2.066287],accel_mss,speed_ms,0,blend_radius_m)
  movel([0.493042, -1.288151, -2.630110, -0.794128, 1.570796, 2.063839],accel_mss,speed_ms,0,blend_radius_m)
  movel([0.491173, -1.287374, -2.630561, -0.794454, 1.570796, 2.061970],accel_mss,speed_ms,0,blend_radius_m)
  movel([0.489831, -1.286234, -2.631221, -0.794934, 1.570796, 2.060627],accel_mss,speed_ms,0,blend_radius_m)
  movel([0.488967, -1.284769, -2.632067, -0.795553, 1.570796, 2.059763],accel_mss,speed_ms,0,blend_radius_m)
  movel([0.488535, -1.283014, -2.633076, -0.796299, 1.570796, 2.059331],accel_mss,speed_ms,0,blend_radius_m)
  movel([0.488483, -1.281012, -2.634224, -0.797154, 1.570796, 2.059279],accel_mss,speed_ms,0,blend_radius_m)
  movel([0.488765, -1.278802, -2.635484, -0.798103, 1.570796, 2.059561],accel_mss,speed_ms,0,blend_radius_m)
  movel([0.489328, -1.276420, -2.636835, -0.799133, 1.570796, 2.060125],accel_mss,speed_ms,0,blend_radius_m)
  movel([0.491106, -1.271321, -2.639705, -0.801363, 1.570796, 2.061903],accel_mss,speed_ms,0,blend_radius_m)
  movel([0.493420, -1.266046, -2.642640, -0.803703, 1.570796, 2.064217],accel_mss,speed_ms,0,blend_radius_m)
  movel([0.497978, -1.256390, -2.647924, -0.808075, 1.570796, 2.068774],accel_mss,speed_ms,0,blend_radius_m)
  movel([0.499662, -1.252124, -2.650223, -0.810043, 1.570796, 2.070458],accel_mss,speed_ms,0,blend_radius_m)
  movel([0.501258, -1.247194, -2.652851, -0.812344, 1.570796, 2.072054],accel_mss,speed_ms,0,blend_radius_m)
  movel([0.502664, -1.241857, -2.655664, -0.814867, 1.570796, 2.073460],accel_mss,speed_ms,0,blend_radius_m)
  movel([0.503778, -1.236372, -2.658521, -0.817496, 1.570796, 2.074575],accel_mss,speed_ms,0,blend_radius_m)
  movel([0.504485, -1.231009, -2.661279, -0.820100, 1.570796, 2.075282],accel_mss,speed_ms,0,blend_radius_m)
  movel([0.504673, -1.226047, -2.663802, -0.822539, 1.570796, 2.075469],accel_mss,speed_ms,0,blend_radius_m)
  movel([0.504225, -1.221778, -2.665950, -0.824661, 1.570796, 2.075021],accel_mss,speed_ms,0,blend_radius_m)
  movel([0.503727, -1.219996, -2.666841, -0.825553, 1.570796, 2.074523],accel_mss,speed_ms,0,blend_radius_m)
  movel([0.503027, -1.218495, -2.667588, -0.826306, 1.570796, 2.073823],accel_mss,speed_ms,0,blend_radius_m)
  movel([0.502054, -1.217160, -2.668250, -0.826979, 1.570796, 2.072850],accel_mss,speed_ms,0,blend_radius_m)
  movel([0.500688, -1.215811, -2.668917, -0.827661, 1.570796, 2.071484],accel_mss,speed_ms,0,blend_radius_m)
  movel([0.498954, -1.214585, -2.669522, -0.828282, 1.570796, 2.069751],accel_mss,speed_ms,0,blend_radius_m)
  movel([0.496884, -1.213620, -2.669997, -0.828772, 1.570796, 2.067681],accel_mss,speed_ms,0,blend_radius_m)
  movel([0.494507, -1.213059, -2.670272, -0.829058, 1.570796, 2.065303],accel_mss,speed_ms,0,blend_radius_m)
  movel([0.491853, -1.213037, -2.670283, -0.829069, 1.570796, 2.062649],accel_mss,speed_ms,0,blend_radius_m)
  movel([0.488959, -1.213692, -2.669961, -0.828735, 1.570796, 2.059755],accel_mss,speed_ms,0,blend_radius_m)
  movel([0.487431, -1.214318, -2.669653, -0.828418, 1.570796, 2.058228],accel_mss,speed_ms,0,blend_radius_m)
  movel([0.485859, -1.215160, -2.669239, -0.827990, 1.570796, 2.056655],accel_mss,speed_ms,0,blend_radius_m)
  movel([0.483530, -1.216849, -2.668404, -0.827136, 1.570796, 2.054326],accel_mss,speed_ms,0,blend_radius_m)
  movel([0.481723, -1.218764, -2.667454, -0.826171, 1.570796, 2.052519],accel_mss,speed_ms,0,blend_radius_m)
  movel([0.480393, -1.220866, -2.666406, -0.825117, 1.570796, 2.051189],accel_mss,speed_ms,0,blend_radius_m)
  movel([0.479488, -1.223120, -2.665277, -0.823992, 1.570796, 2.050284],accel_mss,speed_ms,0,blend_radius_m)
  movel([0.478964, -1.225489, -2.664084, -0.822816, 1.570796, 2.049760],accel_mss,speed_ms,0,blend_radius_m)
  movel([0.478764, -1.227947, -2.662840, -0.821602, 1.570796, 2.049561],accel_mss,speed_ms,0,blend_radius_m)
  movel([0.478841, -1.230456, -2.661562, -0.820371, 1.570796, 2.049637],accel_mss,speed_ms,0,blend_radius_m)
  movel([0.479145, -1.232989, -2.660265, -0.819135, 1.570796, 2.049942],accel_mss,speed_ms,0,blend_radius_m)
  movel([0.480236, -1.237994, -2.657680, -0.816715, 1.570796, 2.051032],accel_mss,speed_ms,0,blend_radius_m)
  movel([0.481654, -1.242716, -2.655214, -0.814459, 1.570796, 2.052450],accel_mss,speed_ms,0,blend_radius_m)
  movel([0.483024, -1.246903, -2.653005, -0.812480, 1.570796, 2.053821],accel_mss,speed_ms,0,blend_radius_m)
  movel([0.483974, -1.250317, -2.651190, -0.810883, 1.570796, 2.054770],accel_mss,speed_ms,0,blend_radius_m)
  movel([0.485853, -1.258763, -2.646636, -0.806990, 1.570796, 2.056649],accel_mss,speed_ms,0,blend_radius_m)
  movel([0.486718, -1.263323, -2.644142, -0.804924, 1.570796, 2.057514],accel_mss,speed_ms,0,blend_radius_m)
  movel([0.487119, -1.267019, -2.642101, -0.803269, 1.570796, 2.057916],accel_mss,speed_ms,0,blend_radius_m)
  movel([0.487043, -1.268572, -2.641239, -0.802578, 1.570796, 2.057839],accel_mss,speed_ms,0,blend_radius_m)
  movel([0.486758, -1.270161, -2.640354, -0.801874, 1.570796, 2.057554],accel_mss,speed_ms,0,blend_radius_m)
  movel([0.485621, -1.273412, -2.638532, -0.800444, 1.570796, 2.056418],accel_mss,speed_ms,0,blend_radius_m)
  movel([0.483836, -1.276681, -2.636688, -0.799020, 1.570796, 2.054633],accel_mss,speed_ms,0,blend_radius_m)
  movel([0.481532, -1.279886, -2.634866, -0.797636, 1.570796, 2.052328],accel_mss,speed_ms,0,blend_radius_m)
  movel([0.478830, -1.282944, -2.633117, -0.796329, 1.570796, 2.049626],accel_mss,speed_ms,0,blend_radius_m)
  movel([0.475850, -1.285774, -2.631487, -0.795128, 1.570796, 2.046647],accel_mss,speed_ms,0,blend_radius_m)
  movel([0.472710, -1.288296, -2.630025, -0.794067, 1.570796, 2.043506],accel_mss,speed_ms,0,blend_radius_m)
  movel([0.469527, -1.290437, -2.628779, -0.793173, 1.570796, 2.040323],accel_mss,speed_ms,0,blend_radius_m)
  movel([0.465555, -1.292552, -2.627542, -0.792295, 1.570796, 2.036351],accel_mss,speed_ms,0,blend_radius_m)
  movel([0.463881, -1.293207, -2.627158, -0.792025, 1.570796, 2.034677],accel_mss,speed_ms,0,blend_radius_m)
  movel([0.462384, -1.293625, -2.626912, -0.791852, 1.570796, 2.033180],accel_mss,speed_ms,0,blend_radius_m)
  movel([0.461042, -1.293827, -2.626793, -0.791769, 1.570796, 2.031838],accel_mss,speed_ms,0,blend_radius_m)
  movel([0.459828, -1.293834, -2.626789, -0.791766, 1.570796, 2.030624],accel_mss,speed_ms,0,blend_radius_m)
  movel([0.457705, -1.293342, -2.627078, -0.791969, 1.570796, 2.028501],accel_mss,speed_ms,0,blend_radius_m)
  movel([0.455831, -1.292322, -2.627676, -0.792390, 1.570796, 2.026628],accel_mss,speed_ms,0,blend_radius_m)
  movel([0.454033, -1.290943, -2.628484, -0.792962, 1.570796, 2.024829],accel_mss,speed_ms,0,blend_radius_m)
  movel([0.449944, -1.287781, -2.630325, -0.794283, 1.570796, 2.020740],accel_mss,speed_ms,0,blend_radius_m)
  movel([0.449705, -1.287647, -2.630402, -0.794339, 1.570796, 2.020501],accel_mss,speed_ms,0,blend_radius_m)
  movel([0.449694, -1.287803, -2.630312, -0.794274, 1.570796, 2.020490],accel_mss,speed_ms,0,blend_radius_m)
  movel([0.450223, -1.288831, -2.629715, -0.793843, 1.570796, 2.021019],accel_mss,speed_ms,0,blend_radius_m)
  movel([0.452693, -1.292674, -2.627470, -0.792245, 1.570796, 2.023489],accel_mss,speed_ms,0,blend_radius_m)
  movel([0.456769, -1.299019, -2.623723, -0.789647, 1.570796, 2.027566],accel_mss,speed_ms,0,blend_radius_m)
  movel([0.452448, -1.297789, -2.624453, -0.790146, 1.570796, 2.023244],accel_mss,speed_ms,0,blend_radius_m)
  movel([0.447836, -1.296123, -2.625440, -0.790826, 1.570796, 2.018632],accel_mss,speed_ms,0,blend_radius_m)
  movel([0.443069, -1.294116, -2.626623, -0.791650, 1.570796, 2.013865],accel_mss,speed_ms,0,blend_radius_m)
  movel([0.438281, -1.291865, -2.627944, -0.792580, 1.570796, 2.009077],accel_mss,speed_ms,0,blend_radius_m)
  movel([0.429221, -1.286975, -2.630792, -0.794622, 1.570796, 2.000017],accel_mss,speed_ms,0,blend_radius_m)
  movel([0.425246, -1.284508, -2.632217, -0.795664, 1.570796, 1.996042],accel_mss,speed_ms,0,blend_radius_m)
  movel([0.421850, -1.282134, -2.633581, -0.796674, 1.570796, 1.992646],accel_mss,speed_ms,0,blend_radius_m)
  movel([0.414634, -1.281863, -2.633736, -0.796789, 1.570796, 1.985430],accel_mss,speed_ms,0,blend_radius_m)
  movel([0.406927, -1.282040, -2.633635, -0.796714, 1.570796, 1.977724],accel_mss,speed_ms,0,blend_radius_m)
  movel([0.390773, -1.283095, -2.633030, -0.796264, 1.570796, 1.961569],accel_mss,speed_ms,0,blend_radius_m)
  movel([0.382673, -1.283655, -2.632708, -0.796026, 1.570796, 1.953470],accel_mss,speed_ms,0,blend_radius_m)
  movel([0.374794, -1.284017, -2.632500, -0.795872, 1.570796, 1.945591],accel_mss,speed_ms,0,blend_radius_m)
  movel([0.367300, -1.284010, -2.632504, -0.795875, 1.570796, 1.938097],accel_mss,speed_ms,0,blend_radius_m)
  movel([0.360355, -1.283466, -2.632817, -0.796106, 1.570796, 1.931152],accel_mss,speed_ms,0,blend_radius_m)
  movel([0.357850, -1.283002, -2.633084, -0.796304, 1.570796, 1.928646],accel_mss,speed_ms,0,blend_radius_m)
  movel([0.355662, -1.282317, -2.633476, -0.796596, 1.570796, 1.926458],accel_mss,speed_ms,0,blend_radius_m)
  movel([0.353797, -1.281422, -2.633989, -0.796978, 1.570796, 1.924594],accel_mss,speed_ms,0,blend_radius_m)
  movel([0.352261, -1.280331, -2.634612, -0.797445, 1.570796, 1.923057],accel_mss,speed_ms,0,blend_radius_m)
  movel([0.351061, -1.279054, -2.635340, -0.797994, 1.570796, 1.921858],accel_mss,speed_ms,0,blend_radius_m)
  movel([0.350202, -1.277607, -2.636163, -0.798619, 1.570796, 1.920998],accel_mss,speed_ms,0,blend_radius_m)
  movel([0.349696, -1.275995, -2.637076, -0.799318, 1.570796, 1.920492],accel_mss,speed_ms,0,blend_radius_m)
  movel([0.349547, -1.274231, -2.638071, -0.800086, 1.570796, 1.920344],accel_mss,speed_ms,0,blend_radius_m)
  movel([0.349765, -1.272334, -2.639138, -0.800917, 1.570796, 1.920561],accel_mss,speed_ms,0,blend_radius_m)
  movel([0.350359, -1.270310, -2.640270, -0.801809, 1.570796, 1.921156],accel_mss,speed_ms,0,blend_radius_m)
  movel([0.351337, -1.268171, -2.641462, -0.802756, 1.570796, 1.922134],accel_mss,speed_ms,0,blend_radius_m)
  movel([0.352707, -1.265935, -2.642701, -0.803752, 1.570796, 1.923503],accel_mss,speed_ms,0,blend_radius_m)
  movel([0.354476, -1.263615, -2.643981, -0.804793, 1.570796, 1.925273],accel_mss,speed_ms,0,blend_radius_m)
  movel([0.356654, -1.261223, -2.645294, -0.805873, 1.570796, 1.927451],accel_mss,speed_ms,0,blend_radius_m)
  movel([0.359250, -1.258777, -2.646628, -0.806984, 1.570796, 1.930047],accel_mss,speed_ms,0,blend_radius_m)
  movel([0.362273, -1.256288, -2.647979, -0.808122, 1.570796, 1.933069],accel_mss,speed_ms,0,blend_radius_m)
  movel([0.362324, -1.258975, -2.646520, -0.806893, 1.570796, 1.933121],accel_mss,speed_ms,0,blend_radius_m)
  movel([0.362441, -1.260235, -2.645833, -0.806320, 1.570796, 1.933237],accel_mss,speed_ms,0,blend_radius_m)
  movel([0.362890, -1.261236, -2.645286, -0.805867, 1.570796, 1.933686],accel_mss,speed_ms,0,blend_radius_m)
  movel([0.363602, -1.261716, -2.645024, -0.805650, 1.570796, 1.934398],accel_mss,speed_ms,0,blend_radius_m)
  movel([0.364729, -1.262021, -2.644857, -0.805512, 1.570796, 1.935526],accel_mss,speed_ms,0,blend_radius_m)
  movel([0.368013, -1.262179, -2.644770, -0.805440, 1.570796, 1.938810],accel_mss,speed_ms,0,blend_radius_m)
  movel([0.372312, -1.261871, -2.644939, -0.805579, 1.570796, 1.943108],accel_mss,speed_ms,0,blend_radius_m)
  movel([0.377205, -1.261246, -2.645281, -0.805862, 1.570796, 1.948001],accel_mss,speed_ms,0,blend_radius_m)
  movel([0.387060, -1.259655, -2.646150, -0.806584, 1.570796, 1.957857],accel_mss,speed_ms,0,blend_radius_m)
  movel([0.394163, -1.258528, -2.646764, -0.807097, 1.570796, 1.964960],accel_mss,speed_ms,0,blend_radius_m)
  movel([0.400035, -1.258102, -2.646995, -0.807292, 1.570796, 1.970831],accel_mss,speed_ms,0,blend_radius_m)
  movel([0.405891, -1.257713, -2.647207, -0.807469, 1.570796, 1.976688],accel_mss,speed_ms,0,blend_radius_m)
  movel([0.399795, -1.251415, -2.650602, -0.810372, 1.570796, 1.970592],accel_mss,speed_ms,0,blend_radius_m)
  movel([0.396859, -1.247865, -2.652495, -0.812029, 1.570796, 1.967655],accel_mss,speed_ms,0,blend_radius_m)
  movel([0.394514, -1.243925, -2.654578, -0.813885, 1.570796, 1.965311],accel_mss,speed_ms,0,blend_radius_m)
  movel([0.393692, -1.241773, -2.655709, -0.814907, 1.570796, 1.964489],accel_mss,speed_ms,0,blend_radius_m)
  movel([0.393169, -1.239479, -2.656907, -0.816002, 1.570796, 1.963965],accel_mss,speed_ms,0,blend_radius_m)
  movel([0.392998, -1.237034, -2.658178, -0.817177, 1.570796, 1.963794],accel_mss,speed_ms,0,blend_radius_m)
  movel([0.393234, -1.234416, -2.659531, -0.818442, 1.570796, 1.964030],accel_mss,speed_ms,0,blend_radius_m)
  movel([0.393927, -1.231614, -2.660970, -0.819805, 1.570796, 1.964723],accel_mss,speed_ms,0,blend_radius_m)
  movel([0.395132, -1.228612, -2.662502, -0.821275, 1.570796, 1.965928],accel_mss,speed_ms,0,blend_radius_m)
  movel([0.396904, -1.225393, -2.664133, -0.822863, 1.570796, 1.967700],accel_mss,speed_ms,0,blend_radius_m)
  movel([0.399300, -1.221945, -2.665866, -0.824577, 1.570796, 1.970097],accel_mss,speed_ms,0,blend_radius_m)
  movel([0.402637, -1.218085, -2.667791, -0.826513, 1.570796, 1.973433],accel_mss,speed_ms,0,blend_radius_m)
  movel([0.406506, -1.214477, -2.669575, -0.828337, 1.570796, 1.977303],accel_mss,speed_ms,0,blend_radius_m)
  movel([0.410763, -1.211220, -2.671173, -0.829996, 1.570796, 1.981559],accel_mss,speed_ms,0,blend_radius_m)
  movel([0.415257, -1.208412, -2.672541, -0.831436, 1.570796, 1.986053],accel_mss,speed_ms,0,blend_radius_m)
  movel([0.419838, -1.206144, -2.673639, -0.832606, 1.570796, 1.990634],accel_mss,speed_ms,0,blend_radius_m)
  movel([0.424353, -1.204521, -2.674422, -0.833446, 1.570796, 1.995149],accel_mss,speed_ms,0,blend_radius_m)
  movel([0.428643, -1.203635, -2.674848, -0.833906, 1.570796, 1.999439],accel_mss,speed_ms,0,blend_radius_m)
  movel([0.432553, -1.203571, -2.674878, -0.833940, 1.570796, 2.003349],accel_mss,speed_ms,0,blend_radius_m)
  movel([0.434271, -1.204156, -2.674597, -0.833636, 1.570796, 2.005067],accel_mss,speed_ms,0,blend_radius_m)
  movel([0.435734, -1.205343, -2.674026, -0.833020, 1.570796, 2.006530],accel_mss,speed_ms,0,blend_radius_m)
  movel([0.436439, -1.206794, -2.673325, -0.832270, 1.570796, 2.007236],accel_mss,speed_ms,0,blend_radius_m)
  movel([0.436352, -1.207516, -2.672975, -0.831898, 1.570796, 2.007148],accel_mss,speed_ms,0,blend_radius_m)
  movel([0.435885, -1.208178, -2.672654, -0.831557, 1.570796, 2.006681],accel_mss,speed_ms,0,blend_radius_m)
  movel([0.434757, -1.207214, -2.673122, -0.832053, 1.570796, 2.005553],accel_mss,speed_ms,0,blend_radius_m)
  movel([0.433605, -1.206606, -2.673416, -0.832367, 1.570796, 2.004401],accel_mss,speed_ms,0,blend_radius_m)
  movel([0.432448, -1.206331, -2.673549, -0.832509, 1.570796, 2.003244],accel_mss,speed_ms,0,blend_radius_m)
  movel([0.431299, -1.206357, -2.673536, -0.832496, 1.570796, 2.002095],accel_mss,speed_ms,0,blend_radius_m)
  movel([0.430170, -1.206660, -2.673390, -0.832339, 1.570796, 2.000967],accel_mss,speed_ms,0,blend_radius_m)
  movel([0.429076, -1.207211, -2.673123, -0.832055, 1.570796, 1.999873],accel_mss,speed_ms,0,blend_radius_m)
  movel([0.428035, -1.207982, -2.672749, -0.831658, 1.570796, 1.998831],accel_mss,speed_ms,0,blend_radius_m)
  movel([0.427061, -1.208941, -2.672284, -0.831164, 1.570796, 1.997858],accel_mss,speed_ms,0,blend_radius_m)
  movel([0.425356, -1.211323, -2.671122, -0.829943, 1.570796, 1.996153],accel_mss,speed_ms,0,blend_radius_m)
  movel([0.424078, -1.214129, -2.669747, -0.828514, 1.570796, 1.994875],accel_mss,speed_ms,0,blend_radius_m)
  movel([0.423320, -1.217145, -2.668257, -0.826986, 1.570796, 1.994116],accel_mss,speed_ms,0,blend_radius_m)
  movel([0.423190, -1.220151, -2.666763, -0.825475, 1.570796, 1.993986],accel_mss,speed_ms,0,blend_radius_m)
  movel([0.423489, -1.221769, -2.665955, -0.824665, 1.570796, 1.994285],accel_mss,speed_ms,0,blend_radius_m)
  movel([0.424134, -1.223528, -2.665072, -0.823789, 1.570796, 1.994930],accel_mss,speed_ms,0,blend_radius_m)
  movel([0.426292, -1.227357, -2.663139, -0.821893, 1.570796, 1.997088],accel_mss,speed_ms,0,blend_radius_m)
  movel([0.429321, -1.231450, -2.661054, -0.819885, 1.570796, 2.000118],accel_mss,speed_ms,0,blend_radius_m)
  movel([0.432884, -1.235604, -2.658918, -0.817867, 1.570796, 2.003680],accel_mss,speed_ms,0,blend_radius_m)
  movel([0.440326, -1.243304, -2.654905, -0.814180, 1.570796, 2.011122],accel_mss,speed_ms,0,blend_radius_m)
  movel([0.446154, -1.248804, -2.651996, -0.811589, 1.570796, 2.016951],accel_mss,speed_ms,0,blend_radius_m)
  movel([0.449097, -1.251531, -2.650540, -0.810318, 1.570796, 2.019893],accel_mss,speed_ms,0,blend_radius_m)
  movel([0.450769, -1.252901, -2.649805, -0.809683, 1.570796, 2.021565],accel_mss,speed_ms,0,blend_radius_m)
  movel([0.452214, -1.253744, -2.649352, -0.809293, 1.570796, 2.023011],accel_mss,speed_ms,0,blend_radius_m)
  movel([0.452721, -1.253843, -2.649299, -0.809247, 1.570796, 2.023518],accel_mss,speed_ms,0,blend_radius_m)
  movel([0.453074, -1.253703, -2.649374, -0.809312, 1.570796, 2.023871],accel_mss,speed_ms,0,blend_radius_m)
  movel([0.453566, -1.252750, -2.649886, -0.809752, 1.570796, 2.024362],accel_mss,speed_ms,0,blend_radius_m)
  movel([0.454197, -1.250006, -2.651356, -0.811028, 1.570796, 2.024993],accel_mss,speed_ms,0,blend_radius_m)
  movel([0.454356, -1.247304, -2.652793, -0.812292, 1.570796, 2.025152],accel_mss,speed_ms,0,blend_radius_m)
  movel([0.454429, -1.241577, -2.655811, -0.815000, 1.570796, 2.025225],accel_mss,speed_ms,0,blend_radius_m)
  movel([0.454940, -1.238326, -2.657507, -0.816555, 1.570796, 2.025737],accel_mss,speed_ms,0,blend_radius_m)
  movel([0.456172, -1.234654, -2.659409, -0.818327, 1.570796, 2.026968],accel_mss,speed_ms,0,blend_radius_m)
  movel([0.457156, -1.232622, -2.660454, -0.819314, 1.570796, 2.027953],accel_mss,speed_ms,0,blend_radius_m)
  movel([0.458440, -1.230437, -2.661572, -0.820380, 1.570796, 2.029237],accel_mss,speed_ms,0,blend_radius_m)
  movel([0.460059, -1.228082, -2.662771, -0.821536, 1.570796, 2.030856],accel_mss,speed_ms,0,blend_radius_m)
  movel([0.462060, -1.225544, -2.664057, -0.822788, 1.570796, 2.032856],accel_mss,speed_ms,0,blend_radius_m)
  movel([0.465013, -1.222378, -2.665650, -0.824362, 1.570796, 2.035809],accel_mss,speed_ms,0,blend_radius_m)
  movel([0.468145, -1.219673, -2.667001, -0.825714, 1.570796, 2.038941],accel_mss,speed_ms,0,blend_radius_m)
  movel([0.471417, -1.217395, -2.668133, -0.826860, 1.570796, 2.042214],accel_mss,speed_ms,0,blend_radius_m)
  movel([0.474793, -1.215508, -2.669067, -0.827814, 1.570796, 2.045589],accel_mss,speed_ms,0,blend_radius_m)
  movel([0.478239, -1.213972, -2.669824, -0.828593, 1.570796, 2.049036],accel_mss,speed_ms,0,blend_radius_m)
  movel([0.481715, -1.212746, -2.670426, -0.829217, 1.570796, 2.052511],accel_mss,speed_ms,0,blend_radius_m)
  movel([0.485189, -1.211787, -2.670895, -0.829706, 1.570796, 2.055986],accel_mss,speed_ms,0,blend_radius_m)
  movel([0.488623, -1.211055, -2.671254, -0.830081, 1.570796, 2.059419],accel_mss,speed_ms,0,blend_radius_m)
  movel([0.494812, -1.210302, -2.671621, -0.830466, 1.570796, 2.065608],accel_mss,speed_ms,0,blend_radius_m)
  movel([0.499838, -1.210382, -2.671582, -0.830425, 1.570796, 2.070634],accel_mss,speed_ms,0,blend_radius_m)
  movel([0.503701, -1.211002, -2.671279, -0.830108, 1.570796, 2.074498],accel_mss,speed_ms,0,blend_radius_m)
  movel([0.506413, -1.211859, -2.670860, -0.829670, 1.570796, 2.077209],accel_mss,speed_ms,0,blend_radius_m)
  movel([0.509892, -1.213781, -2.669917, -0.828690, 1.570796, 2.080688],accel_mss,speed_ms,0,blend_radius_m)
  movel([0.512653, -1.216339, -2.668656, -0.827394, 1.570796, 2.083449],accel_mss,speed_ms,0,blend_radius_m)
  movel([0.514710, -1.219455, -2.667110, -0.825824, 1.570796, 2.085506],accel_mss,speed_ms,0,blend_radius_m)
  movel([0.516075, -1.223050, -2.665313, -0.824027, 1.570796, 2.086871],accel_mss,speed_ms,0,blend_radius_m)
  movel([0.516761, -1.227041, -2.663299, -0.822048, 1.570796, 2.087557],accel_mss,speed_ms,0,blend_radius_m)
  movel([0.516786, -1.231353, -2.661104, -0.819932, 1.570796, 2.087582],accel_mss,speed_ms,0,blend_radius_m)
  movel([0.516164, -1.235915, -2.658757, -0.817717, 1.570796, 2.086960],accel_mss,speed_ms,0,blend_radius_m)
  movel([0.514913, -1.240652, -2.656295, -0.815442, 1.570796, 2.085709],accel_mss,speed_ms,0,blend_radius_m)
  movel([0.513258, -1.245009, -2.654007, -0.813373, 1.570796, 2.084055],accel_mss,speed_ms,0,blend_radius_m)
  movel([0.511317, -1.249348, -2.651706, -0.811335, 1.570796, 2.082113],accel_mss,speed_ms,0,blend_radius_m)
  movel([0.509367, -1.253599, -2.649430, -0.809360, 1.570796, 2.080163],accel_mss,speed_ms,0,blend_radius_m)
  movel([0.507692, -1.257701, -2.647213, -0.807475, 1.570796, 2.078489],accel_mss,speed_ms,0,blend_radius_m)
  movel([0.506568, -1.261580, -2.645098, -0.805711, 1.570796, 2.077364],accel_mss,speed_ms,0,blend_radius_m)
  movel([0.506296, -1.263417, -2.644090, -0.804882, 1.570796, 2.077093],accel_mss,speed_ms,0,blend_radius_m)
  movel([0.506263, -1.265178, -2.643120, -0.804091, 1.570796, 2.077060],accel_mss,speed_ms,0,blend_radius_m)
  movel([0.506504, -1.266852, -2.642194, -0.803343, 1.570796, 2.077301],accel_mss,speed_ms,0,blend_radius_m)
  movel([0.507050, -1.268435, -2.641315, -0.802639, 1.570796, 2.077847],accel_mss,speed_ms,0,blend_radius_m)
  movel([0.507932, -1.269918, -2.640489, -0.801982, 1.570796, 2.078728],accel_mss,speed_ms,0,blend_radius_m)
  movel([0.509186, -1.271297, -2.639719, -0.801373, 1.570796, 2.079982],accel_mss,speed_ms,0,blend_radius_m)
  movel([0.510577, -1.272215, -2.639204, -0.800970, 1.570796, 2.081374],accel_mss,speed_ms,0,blend_radius_m)
  movel([0.512099, -1.272613, -2.638981, -0.800795, 1.570796, 2.082895],accel_mss,speed_ms,0,blend_radius_m)
  movel([0.513705, -1.272557, -2.639012, -0.800819, 1.570796, 2.084502],accel_mss,speed_ms,0,blend_radius_m)
  movel([0.515345, -1.272107, -2.639265, -0.801017, 1.570796, 2.086142],accel_mss,speed_ms,0,blend_radius_m)
  movel([0.516975, -1.271323, -2.639704, -0.801362, 1.570796, 2.087771],accel_mss,speed_ms,0,blend_radius_m)
  movel([0.518542, -1.270270, -2.640293, -0.801826, 1.570796, 2.089338],accel_mss,speed_ms,0,blend_radius_m)
  movel([0.519999, -1.269004, -2.640999, -0.802387, 1.570796, 2.090796],accel_mss,speed_ms,0,blend_radius_m)
  movel([0.521296, -1.267586, -2.641787, -0.803016, 1.570796, 2.092092],accel_mss,speed_ms,0,blend_radius_m)
  movel([0.522382, -1.266082, -2.642620, -0.803687, 1.570796, 2.093178],accel_mss,speed_ms,0,blend_radius_m)
  movel([0.523206, -1.264548, -2.643467, -0.804374, 1.570796, 2.094003],accel_mss,speed_ms,0,blend_radius_m)
  movel([0.523716, -1.263052, -2.644290, -0.805046, 1.570796, 2.094512],accel_mss,speed_ms,0,blend_radius_m)
  movel([0.523860, -1.261653, -2.645058, -0.805678, 1.570796, 2.094656],accel_mss,speed_ms,0,blend_radius_m)
  movel([0.523580, -1.260421, -2.645732, -0.806236, 1.570796, 2.094376],accel_mss,speed_ms,0,blend_radius_m)
  movel([0.522828, -1.259420, -2.646278, -0.806691, 1.570796, 2.093624],accel_mss,speed_ms,0,blend_radius_m)
  movel([0.521552, -1.258714, -2.646663, -0.807013, 1.570796, 2.092348],accel_mss,speed_ms,0,blend_radius_m)
  movel([0.519693, -1.258374, -2.646847, -0.807167, 1.570796, 2.090490],accel_mss,speed_ms,0,blend_radius_m)
  movel([0.519939, -1.259561, -2.646202, -0.806627, 1.570796, 2.090735],accel_mss,speed_ms,0,blend_radius_m)
  movel([0.519863, -1.260723, -2.645567, -0.806099, 1.570796, 2.090659],accel_mss,speed_ms,0,blend_radius_m)
  movel([0.519492, -1.261825, -2.644964, -0.805600, 1.570796, 2.090289],accel_mss,speed_ms,0,blend_radius_m)
  movel([0.518855, -1.262817, -2.644420, -0.805152, 1.570796, 2.089651],accel_mss,speed_ms,0,blend_radius_m)
  movel([0.517973, -1.263669, -2.643951, -0.804769, 1.570796, 2.088770],accel_mss,speed_ms,0,blend_radius_m)
  movel([0.516879, -1.264335, -2.643584, -0.804469, 1.570796, 2.087676],accel_mss,speed_ms,0,blend_radius_m)
  movel([0.515591, -1.264776, -2.643342, -0.804272, 1.570796, 2.086387],accel_mss,speed_ms,0,blend_radius_m)
  movel([0.514135, -1.264957, -2.643242, -0.804190, 1.570796, 2.084932],accel_mss,speed_ms,0,blend_radius_m)
  movel([0.511917, -1.264685, -2.643391, -0.804312, 1.570796, 2.082714],accel_mss,speed_ms,0,blend_radius_m)
  movel([0.510374, -1.263815, -2.643871, -0.804703, 1.570796, 2.081170],accel_mss,speed_ms,0,blend_radius_m)
  movel([0.509457, -1.262426, -2.644634, -0.805329, 1.570796, 2.080253],accel_mss,speed_ms,0,blend_radius_m)
  movel([0.509120, -1.260612, -2.645627, -0.806149, 1.570796, 2.079916],accel_mss,speed_ms,0,blend_radius_m)
  movel([0.509319, -1.258452, -2.646805, -0.807132, 1.570796, 2.080115],accel_mss,speed_ms,0,blend_radius_m)
  movel([0.510008, -1.256038, -2.648114, -0.808237, 1.570796, 2.080804],accel_mss,speed_ms,0,blend_radius_m)
  movel([0.511145, -1.253453, -2.649509, -0.809427, 1.570796, 2.081942],accel_mss,speed_ms,0,blend_radius_m)
  movel([0.512682, -1.250794, -2.650934, -0.810660, 1.570796, 2.083478],accel_mss,speed_ms,0,blend_radius_m)
  movel([0.514578, -1.248148, -2.652345, -0.811896, 1.570796, 2.085374],accel_mss,speed_ms,0,blend_radius_m)
  movel([0.516781, -1.245612, -2.653689, -0.813088, 1.570796, 2.087577],accel_mss,speed_ms,0,blend_radius_m)
  movel([0.519243, -1.243280, -2.654918, -0.814191, 1.570796, 2.090039],accel_mss,speed_ms,0,blend_radius_m)
  movel([0.521912, -1.241254, -2.655981, -0.815155, 1.570796, 2.092709],accel_mss,speed_ms,0,blend_radius_m)
  movel([0.524738, -1.239632, -2.656828, -0.815929, 1.570796, 2.095534],accel_mss,speed_ms,0,blend_radius_m)
  movel([0.527663, -1.238513, -2.657410, -0.816466, 1.570796, 2.098459],accel_mss,speed_ms,0,blend_radius_m)
  movel([0.530635, -1.237996, -2.657679, -0.816714, 1.570796, 2.101431],accel_mss,speed_ms,0,blend_radius_m)
  movel([0.533592, -1.238182, -2.657582, -0.816625, 1.570796, 2.104389],accel_mss,speed_ms,0,blend_radius_m)
  movel([0.535510, -1.238688, -2.657319, -0.816382, 1.570796, 2.106306],accel_mss,speed_ms,0,blend_radius_m)
  movel([0.537243, -1.239415, -2.656941, -0.816033, 1.570796, 2.108039],accel_mss,speed_ms,0,blend_radius_m)
  movel([0.538782, -1.240352, -2.656452, -0.815585, 1.570796, 2.109579],accel_mss,speed_ms,0,blend_radius_m)
  movel([0.540118, -1.241482, -2.655861, -0.815046, 1.570796, 2.110914],accel_mss,speed_ms,0,blend_radius_m)
  movel([0.541244, -1.242795, -2.655173, -0.814421, 1.570796, 2.112041],accel_mss,speed_ms,0,blend_radius_m)
  movel([0.542156, -1.244276, -2.654394, -0.813720, 1.570796, 2.112952],accel_mss,speed_ms,0,blend_radius_m)
  movel([0.542841, -1.245906, -2.653533, -0.812950, 1.570796, 2.113637],accel_mss,speed_ms,0,blend_radius_m)
  movel([0.543297, -1.247676, -2.652595, -0.812117, 1.570796, 2.114094],accel_mss,speed_ms,0,blend_radius_m)
  movel([0.543513, -1.249571, -2.651588, -0.811231, 1.570796, 2.114309],accel_mss,speed_ms,0,blend_radius_m)
  movel([0.543487, -1.251576, -2.650516, -0.810297, 1.570796, 2.114283],accel_mss,speed_ms,0,blend_radius_m)
  movel([0.543210, -1.253677, -2.649388, -0.809324, 1.570796, 2.114007],accel_mss,speed_ms,0,blend_radius_m)
  movel([0.542681, -1.255861, -2.648210, -0.808318, 1.570796, 2.113477],accel_mss,speed_ms,0,blend_radius_m)
  movel([0.541885, -1.258117, -2.646987, -0.807285, 1.570796, 2.112681],accel_mss,speed_ms,0,blend_radius_m)
  movel([0.540822, -1.260429, -2.645728, -0.806232, 1.570796, 2.111618],accel_mss,speed_ms,0,blend_radius_m)
  movel([0.539486, -1.262787, -2.644436, -0.805166, 1.570796, 2.110282],accel_mss,speed_ms,0,blend_radius_m)
  movel([0.537867, -1.265178, -2.643120, -0.804091, 1.570796, 2.108664],accel_mss,speed_ms,0,blend_radius_m)
  movel([0.535863, -1.267386, -2.641898, -0.803105, 1.570796, 2.106659],accel_mss,speed_ms,0,blend_radius_m)
  movel([0.533409, -1.269582, -2.640676, -0.802130, 1.570796, 2.104206],accel_mss,speed_ms,0,blend_radius_m)
  movel([0.531231, -1.271409, -2.639656, -0.801324, 1.570796, 2.102027],accel_mss,speed_ms,0,blend_radius_m)
  movel([0.530051, -1.272511, -2.639039, -0.800840, 1.570796, 2.100847],accel_mss,speed_ms,0,blend_radius_m)
  movel([0.529727, -1.273571, -2.638443, -0.800375, 1.570796, 2.100523],accel_mss,speed_ms,0,blend_radius_m)
  movel([0.529546, -1.275222, -2.637513, -0.799654, 1.570796, 2.100342],accel_mss,speed_ms,0,blend_radius_m)
  movel([0.529353, -1.277036, -2.636487, -0.798866, 1.570796, 2.100149],accel_mss,speed_ms,0,blend_radius_m)
  movel([0.528990, -1.278591, -2.635604, -0.798194, 1.570796, 2.099787],accel_mss,speed_ms,0,blend_radius_m)
  movel([0.528030, -1.280692, -2.634406, -0.797291, 1.570796, 2.098826],accel_mss,speed_ms,0,blend_radius_m)
  movel([0.526853, -1.282644, -2.633289, -0.796456, 1.570796, 2.097649],accel_mss,speed_ms,0,blend_radius_m)
  movel([0.525488, -1.284446, -2.632253, -0.795690, 1.570796, 2.096284],accel_mss,speed_ms,0,blend_radius_m)
  movel([0.523966, -1.286084, -2.631308, -0.794998, 1.570796, 2.094763],accel_mss,speed_ms,0,blend_radius_m)
  movel([0.522314, -1.287554, -2.630456, -0.794379, 1.570796, 2.093110],accel_mss,speed_ms,0,blend_radius_m)
  movel([0.520558, -1.288850, -2.629704, -0.793835, 1.570796, 2.091354],accel_mss,speed_ms,0,blend_radius_m)
  movel([0.518728, -1.289961, -2.629057, -0.793371, 1.570796, 2.089524],accel_mss,speed_ms,0,blend_radius_m)
  movel([0.516850, -1.290885, -2.628517, -0.792986, 1.570796, 2.087646],accel_mss,speed_ms,0,blend_radius_m)
  movel([0.514949, -1.291611, -2.628093, -0.792685, 1.570796, 2.085745],accel_mss,speed_ms,0,blend_radius_m)
  movel([0.513056, -1.292132, -2.627788, -0.792469, 1.570796, 2.083852],accel_mss,speed_ms,0,blend_radius_m)
  movel([0.511194, -1.292438, -2.627609, -0.792342, 1.570796, 2.081990],accel_mss,speed_ms,0,blend_radius_m)
  speed_ms = 0.003
  movel([0.511194, -1.285477, -2.624306, -0.802605, 1.570796, 2.081990],accel_mss,speed_ms,0,blend_radius_m)
  speed_ms = 0.03
  movel([0.511194, -1.258845, -2.610818, -0.842726, 1.570796, 2.081990],accel_mss,speed_ms,0,blend_radius_m)
  #M_RunCode9
  movel([0.516540, -1.266690, -2.606395, -0.839304, 1.570796, 2.087337],accel_mss,speed_ms,0,blend_radius_m)
  #M_RunCode3
  movel([0.516540, -1.293212, -2.619779, -0.799397, 1.570796, 2.087337],accel_mss,speed_ms,0,blend_radius_m)
  speed_ms = 0.003
  movel([0.516540, -1.300140, -2.623056, -0.789193, 1.570796, 2.087337],accel_mss,speed_ms,0,blend_radius_m)
  speed_ms = 0.007
  movel([0.517996, -1.299036, -2.623713, -0.789640, 1.570796, 2.088792],accel_mss,speed_ms,0,blend_radius_m)
  movel([0.521110, -1.297088, -2.624869, -0.790432, 1.570796, 2.091906],accel_mss,speed_ms,0,blend_radius_m)
  movel([0.524092, -1.295089, -2.626050, -0.791250, 1.570796, 2.094889],accel_mss,speed_ms,0,blend_radius_m)
  movel([0.525380, -1.293920, -2.626738, -0.791731, 1.570796, 2.096176],accel_mss,speed_ms,0,blend_radius_m)
  movel([0.526455, -1.292554, -2.627541, -0.792294, 1.570796, 2.097251],accel_mss,speed_ms,0,blend_radius_m)
  movel([0.525946, -1.293622, -2.626914, -0.791853, 1.570796, 2.096743],accel_mss,speed_ms,0,blend_radius_m)
  movel([0.524714, -1.295501, -2.625807, -0.791081, 1.570796, 2.095510],accel_mss,speed_ms,0,blend_radius_m)
  movel([0.523266, -1.297085, -2.624871, -0.790433, 1.570796, 2.094062],accel_mss,speed_ms,0,blend_radius_m)
  movel([0.521662, -1.298475, -2.624046, -0.789868, 1.570796, 2.092458],accel_mss,speed_ms,0,blend_radius_m)
  movel([0.519973, -1.299756, -2.623284, -0.789349, 1.570796, 2.090770],accel_mss,speed_ms,0,blend_radius_m)
  movel([0.516594, -1.302364, -2.621727, -0.788299, 1.570796, 2.087390],accel_mss,speed_ms,0,blend_radius_m)
  movel([0.515039, -1.303871, -2.620822, -0.787696, 1.570796, 2.085835],accel_mss,speed_ms,0,blend_radius_m)
  movel([0.513664, -1.305628, -2.619765, -0.786997, 1.570796, 2.084460],accel_mss,speed_ms,0,blend_radius_m)
  movel([0.512429, -1.307715, -2.618502, -0.786171, 1.570796, 2.083225],accel_mss,speed_ms,0,blend_radius_m)
  movel([0.511858, -1.308843, -2.617818, -0.785727, 1.570796, 2.082655],accel_mss,speed_ms,0,blend_radius_m)
  movel([0.511665, -1.309499, -2.617420, -0.785470, 1.570796, 2.082461],accel_mss,speed_ms,0,blend_radius_m)
  movel([0.512378, -1.309836, -2.617214, -0.785338, 1.570796, 2.083175],accel_mss,speed_ms,0,blend_radius_m)
  movel([0.512930, -1.310152, -2.617022, -0.785215, 1.570796, 2.083726],accel_mss,speed_ms,0,blend_radius_m)
  movel([0.513357, -1.310622, -2.616736, -0.785031, 1.570796, 2.084153],accel_mss,speed_ms,0,blend_radius_m)
  movel([0.513840, -1.311842, -2.615991, -0.784556, 1.570796, 2.084637],accel_mss,speed_ms,0,blend_radius_m)
  movel([0.513949, -1.312926, -2.615327, -0.784136, 1.570796, 2.084745],accel_mss,speed_ms,0,blend_radius_m)
  movel([0.513748, -1.313922, -2.614716, -0.783751, 1.570796, 2.084544],accel_mss,speed_ms,0,blend_radius_m)
  movel([0.513308, -1.314880, -2.614127, -0.783382, 1.570796, 2.084104],accel_mss,speed_ms,0,blend_radius_m)
  movel([0.511974, -1.316871, -2.612899, -0.782618, 1.570796, 2.082770],accel_mss,speed_ms,0,blend_radius_m)
  movel([0.510474, -1.319287, -2.611403, -0.781700, 1.570796, 2.081271],accel_mss,speed_ms,0,blend_radius_m)
  movel([0.508931, -1.322594, -2.609341, -0.780454, 1.570796, 2.079728],accel_mss,speed_ms,0,blend_radius_m)
  movel([0.507517, -1.325877, -2.607280, -0.779232, 1.570796, 2.078313],accel_mss,speed_ms,0,blend_radius_m)
  movel([0.505977, -1.329137, -2.605219, -0.778033, 1.570796, 2.076774],accel_mss,speed_ms,0,blend_radius_m)
  movel([0.504070, -1.332367, -2.603163, -0.776860, 1.570796, 2.074866],accel_mss,speed_ms,0,blend_radius_m)
  movel([0.502813, -1.334060, -2.602079, -0.776250, 1.570796, 2.073609],accel_mss,speed_ms,0,blend_radius_m)
  movel([0.501417, -1.335684, -2.601036, -0.775669, 1.570796, 2.072213],accel_mss,speed_ms,0,blend_radius_m)
  movel([0.498370, -1.338767, -2.599047, -0.774576, 1.570796, 2.069166],accel_mss,speed_ms,0,blend_radius_m)
  movel([0.495231, -1.341716, -2.597131, -0.773542, 1.570796, 2.066027],accel_mss,speed_ms,0,blend_radius_m)
  movel([0.492314, -1.344624, -2.595231, -0.772534, 1.570796, 2.063110],accel_mss,speed_ms,0,blend_radius_m)
  movel([0.487958, -1.349701, -2.591885, -0.770803, 1.570796, 2.058754],accel_mss,speed_ms,0,blend_radius_m)
  movel([0.486144, -1.351890, -2.590431, -0.770068, 1.570796, 2.056940],accel_mss,speed_ms,0,blend_radius_m)
  movel([0.484335, -1.353898, -2.589092, -0.769399, 1.570796, 2.055131],accel_mss,speed_ms,0,blend_radius_m)
  movel([0.482356, -1.355759, -2.587846, -0.768784, 1.570796, 2.053153],accel_mss,speed_ms,0,blend_radius_m)
  movel([0.480031, -1.357514, -2.586667, -0.768209, 1.570796, 2.050827],accel_mss,speed_ms,0,blend_radius_m)
  movel([0.477183, -1.359199, -2.585530, -0.767660, 1.570796, 2.047979],accel_mss,speed_ms,0,blend_radius_m)
  movel([0.473638, -1.360856, -2.584408, -0.767125, 1.570796, 2.044434],accel_mss,speed_ms,0,blend_radius_m)
  movel([0.470735, -1.361947, -2.583668, -0.766774, 1.570796, 2.041531],accel_mss,speed_ms,0,blend_radius_m)
  movel([0.468083, -1.362689, -2.583163, -0.766537, 1.570796, 2.038879],accel_mss,speed_ms,0,blend_radius_m)
  movel([0.465663, -1.363105, -2.582879, -0.766404, 1.570796, 2.036459],accel_mss,speed_ms,0,blend_radius_m)
  movel([0.463467, -1.363219, -2.582802, -0.766368, 1.570796, 2.034263],accel_mss,speed_ms,0,blend_radius_m)
  movel([0.461485, -1.363042, -2.582922, -0.766424, 1.570796, 2.032281],accel_mss,speed_ms,0,blend_radius_m)
  movel([0.459708, -1.362600, -2.583224, -0.766565, 1.570796, 2.030504],accel_mss,speed_ms,0,blend_radius_m)
  movel([0.458120, -1.361908, -2.583694, -0.766787, 1.570796, 2.028916],accel_mss,speed_ms,0,blend_radius_m)
  movel([0.456715, -1.360985, -2.584321, -0.767083, 1.570796, 2.027511],accel_mss,speed_ms,0,blend_radius_m)
  movel([0.455485, -1.359853, -2.585088, -0.767448, 1.570796, 2.026281],accel_mss,speed_ms,0,blend_radius_m)
  movel([0.454417, -1.358528, -2.585983, -0.767878, 1.570796, 2.025213],accel_mss,speed_ms,0,blend_radius_m)
  movel([0.452739, -1.355375, -2.588104, -0.768911, 1.570796, 2.023535],accel_mss,speed_ms,0,blend_radius_m)
  movel([0.451613, -1.351672, -2.590576, -0.770140, 1.570796, 2.022409],accel_mss,speed_ms,0,blend_radius_m)
  movel([0.450973, -1.347572, -2.593292, -0.771525, 1.570796, 2.021769],accel_mss,speed_ms,0,blend_radius_m)
  movel([0.450820, -1.343466, -2.595989, -0.772934, 1.570796, 2.021616],accel_mss,speed_ms,0,blend_radius_m)
  movel([0.450750, -1.338117, -2.599467, -0.774805, 1.570796, 2.021547],accel_mss,speed_ms,0,blend_radius_m)
  movel([0.450379, -1.332284, -2.603216, -0.776890, 1.570796, 2.021176],accel_mss,speed_ms,0,blend_radius_m)
  movel([0.449959, -1.329425, -2.605036, -0.777928, 1.570796, 2.020755],accel_mss,speed_ms,0,blend_radius_m)
  movel([0.449314, -1.326744, -2.606733, -0.778912, 1.570796, 2.020110],accel_mss,speed_ms,0,blend_radius_m)
  movel([0.448394, -1.324341, -2.608246, -0.779802, 1.570796, 2.019190],accel_mss,speed_ms,0,blend_radius_m)
  movel([0.447150, -1.322317, -2.609514, -0.780558, 1.570796, 2.017946],accel_mss,speed_ms,0,blend_radius_m)
  movel([0.445532, -1.320780, -2.610474, -0.781136, 1.570796, 2.016328],accel_mss,speed_ms,0,blend_radius_m)
  movel([0.443493, -1.319831, -2.611064, -0.781494, 1.570796, 2.014289],accel_mss,speed_ms,0,blend_radius_m)
  movel([0.442297, -1.319614, -2.611199, -0.781576, 1.570796, 2.013094],accel_mss,speed_ms,0,blend_radius_m)
  movel([0.440982, -1.319581, -2.611220, -0.781588, 1.570796, 2.011778],accel_mss,speed_ms,0,blend_radius_m)
  movel([0.439536, -1.319749, -2.611115, -0.781525, 1.570796, 2.010332],accel_mss,speed_ms,0,blend_radius_m)
  movel([0.437960, -1.320127, -2.610880, -0.781382, 1.570796, 2.008756],accel_mss,speed_ms,0,blend_radius_m)
  movel([0.436244, -1.320730, -2.610505, -0.781154, 1.570796, 2.007040],accel_mss,speed_ms,0,blend_radius_m)
  movel([0.434386, -1.321568, -2.609982, -0.780839, 1.570796, 2.005183],accel_mss,speed_ms,0,blend_radius_m)
  movel([0.430224, -1.324001, -2.608459, -0.779929, 1.570796, 2.001020],accel_mss,speed_ms,0,blend_radius_m)
  movel([0.428397, -1.325535, -2.607495, -0.779359, 1.570796, 1.999193],accel_mss,speed_ms,0,blend_radius_m)
  movel([0.426728, -1.327309, -2.606376, -0.778704, 1.570796, 1.997525],accel_mss,speed_ms,0,blend_radius_m)
  movel([0.425250, -1.329318, -2.605104, -0.777967, 1.570796, 1.996046],accel_mss,speed_ms,0,blend_radius_m)
  movel([0.423993, -1.331552, -2.603683, -0.777155, 1.570796, 1.994790],accel_mss,speed_ms,0,blend_radius_m)
  movel([0.426796, -1.330448, -2.604386, -0.777555, 1.570796, 1.997592],accel_mss,speed_ms,0,blend_radius_m)
  movel([0.429485, -1.329653, -2.604891, -0.777845, 1.570796, 2.000282],accel_mss,speed_ms,0,blend_radius_m)
  movel([0.432046, -1.329158, -2.605206, -0.778026, 1.570796, 2.002843],accel_mss,speed_ms,0,blend_radius_m)
  movel([0.434463, -1.328957, -2.605333, -0.778099, 1.570796, 2.005259],accel_mss,speed_ms,0,blend_radius_m)
  movel([0.436717, -1.329041, -2.605280, -0.778069, 1.570796, 2.007513],accel_mss,speed_ms,0,blend_radius_m)
  movel([0.438797, -1.329397, -2.605053, -0.777938, 1.570796, 2.009593],accel_mss,speed_ms,0,blend_radius_m)
  movel([0.440681, -1.330022, -2.604656, -0.777710, 1.570796, 2.011477],accel_mss,speed_ms,0,blend_radius_m)
  movel([0.442359, -1.330900, -2.604098, -0.777391, 1.570796, 2.013155],accel_mss,speed_ms,0,blend_radius_m)
  movel([0.443811, -1.332026, -2.603380, -0.776983, 1.570796, 2.014608],accel_mss,speed_ms,0,blend_radius_m)
  movel([0.445031, -1.333383, -2.602513, -0.776493, 1.570796, 2.015828],accel_mss,speed_ms,0,blend_radius_m)
  movel([0.446002, -1.334961, -2.601501, -0.775927, 1.570796, 2.016798],accel_mss,speed_ms,0,blend_radius_m)
  movel([0.446709, -1.336751, -2.600349, -0.775289, 1.570796, 2.017506],accel_mss,speed_ms,0,blend_radius_m)
  movel([0.447142, -1.338740, -2.599064, -0.774585, 1.570796, 2.017938],accel_mss,speed_ms,0,blend_radius_m)
  movel([0.447287, -1.340917, -2.597651, -0.773821, 1.570796, 2.018083],accel_mss,speed_ms,0,blend_radius_m)
  movel([0.447133, -1.343269, -2.596117, -0.773002, 1.570796, 2.017929],accel_mss,speed_ms,0,blend_radius_m)
  movel([0.446672, -1.345787, -2.594467, -0.772134, 1.570796, 2.017468],accel_mss,speed_ms,0,blend_radius_m)
  movel([0.446063, -1.347913, -2.593067, -0.771409, 1.570796, 2.016859],accel_mss,speed_ms,0,blend_radius_m)
  movel([0.445275, -1.349989, -2.591694, -0.770706, 1.570796, 2.016071],accel_mss,speed_ms,0,blend_radius_m)
  movel([0.444321, -1.352009, -2.590352, -0.770028, 1.570796, 2.015118],accel_mss,speed_ms,0,blend_radius_m)
  movel([0.443220, -1.353965, -2.589047, -0.769377, 1.570796, 2.014016],accel_mss,speed_ms,0,blend_radius_m)
  movel([0.440619, -1.357669, -2.586562, -0.768158, 1.570796, 2.011415],accel_mss,speed_ms,0,blend_radius_m)
  movel([0.437580, -1.361054, -2.584274, -0.767061, 1.570796, 2.008377],accel_mss,speed_ms,0,blend_radius_m)
  movel([0.434212, -1.364076, -2.582218, -0.766095, 1.570796, 2.005008],accel_mss,speed_ms,0,blend_radius_m)
  movel([0.430619, -1.366689, -2.580429, -0.765271, 1.570796, 2.001415],accel_mss,speed_ms,0,blend_radius_m)
  movel([0.426897, -1.368854, -2.578940, -0.764595, 1.570796, 1.997693],accel_mss,speed_ms,0,blend_radius_m)
  movel([0.423149, -1.370520, -2.577789, -0.764079, 1.570796, 1.993945],accel_mss,speed_ms,0,blend_radius_m)
  movel([0.419471, -1.371644, -2.577011, -0.763734, 1.570796, 1.990268],accel_mss,speed_ms,0,blend_radius_m)
  movel([0.415963, -1.372179, -2.576640, -0.763570, 1.570796, 1.986760],accel_mss,speed_ms,0,blend_radius_m)
  movel([0.412722, -1.372072, -2.576715, -0.763602, 1.570796, 1.983518],accel_mss,speed_ms,0,blend_radius_m)
  movel([0.411230, -1.371763, -2.576929, -0.763697, 1.570796, 1.982027],accel_mss,speed_ms,0,blend_radius_m)
  movel([0.409843, -1.371272, -2.577270, -0.763848, 1.570796, 1.980640],accel_mss,speed_ms,0,blend_radius_m)
  movel([0.408571, -1.370595, -2.577738, -0.764056, 1.570796, 1.979367],accel_mss,speed_ms,0,blend_radius_m)
  movel([0.407429, -1.369721, -2.578342, -0.764326, 1.570796, 1.978225],accel_mss,speed_ms,0,blend_radius_m)
  movel([0.406427, -1.368643, -2.579086, -0.764661, 1.570796, 1.977223],accel_mss,speed_ms,0,blend_radius_m)
  movel([0.405580, -1.367355, -2.579972, -0.765062, 1.570796, 1.976376],accel_mss,speed_ms,0,blend_radius_m)
  movel([0.404901, -1.365850, -2.581005, -0.765535, 1.570796, 1.975697],accel_mss,speed_ms,0,blend_radius_m)
  movel([0.404405, -1.364114, -2.582191, -0.766083, 1.570796, 1.975201],accel_mss,speed_ms,0,blend_radius_m)
  movel([0.404103, -1.362142, -2.583535, -0.766712, 1.570796, 1.974899],accel_mss,speed_ms,0,blend_radius_m)
  movel([0.404012, -1.359924, -2.585040, -0.767425, 1.570796, 1.974808],accel_mss,speed_ms,0,blend_radius_m)
  movel([0.404253, -1.357992, -2.586345, -0.768053, 1.570796, 1.975050],accel_mss,speed_ms,0,blend_radius_m)
  movel([0.405428, -1.352478, -2.590040, -0.769871, 1.570796, 1.976224],accel_mss,speed_ms,0,blend_radius_m)
  movel([0.406583, -1.348498, -2.592681, -0.771210, 1.570796, 1.977380],accel_mss,speed_ms,0,blend_radius_m)
  movel([0.408235, -1.343765, -2.595793, -0.772831, 1.570796, 1.979031],accel_mss,speed_ms,0,blend_radius_m)
  movel([0.410486, -1.338317, -2.599338, -0.774734, 1.570796, 1.981282],accel_mss,speed_ms,0,blend_radius_m)
  movel([0.413427, -1.332200, -2.603269, -0.776920, 1.570796, 1.984223],accel_mss,speed_ms,0,blend_radius_m)
  movel([0.415823, -1.327898, -2.606004, -0.778487, 1.570796, 1.986620],accel_mss,speed_ms,0,blend_radius_m)
  movel([0.418324, -1.324024, -2.608445, -0.779920, 1.570796, 1.989120],accel_mss,speed_ms,0,blend_radius_m)
  movel([0.420890, -1.320561, -2.610610, -0.781218, 1.570796, 1.991687],accel_mss,speed_ms,0,blend_radius_m)
  movel([0.423488, -1.317493, -2.612515, -0.782381, 1.570796, 1.994284],accel_mss,speed_ms,0,blend_radius_m)
  movel([0.426079, -1.314804, -2.614174, -0.783411, 1.570796, 1.996876],accel_mss,speed_ms,0,blend_radius_m)
  movel([0.428629, -1.312471, -2.615606, -0.784312, 1.570796, 1.999426],accel_mss,speed_ms,0,blend_radius_m)
  movel([0.431102, -1.310473, -2.616826, -0.785089, 1.570796, 2.001898],accel_mss,speed_ms,0,blend_radius_m)
  movel([0.433460, -1.308793, -2.617849, -0.785747, 1.570796, 2.004257],accel_mss,speed_ms,0,blend_radius_m)
  movel([0.437692, -1.306280, -2.619371, -0.786738, 1.570796, 2.008488],accel_mss,speed_ms,0,blend_radius_m)
  movel([0.441048, -1.304744, -2.620297, -0.787348, 1.570796, 2.011844],accel_mss,speed_ms,0,blend_radius_m)
  movel([0.443252, -1.303977, -2.620759, -0.787653, 1.570796, 2.014048],accel_mss,speed_ms,0,blend_radius_m)
  movel([0.444045, -1.303768, -2.620884, -0.787737, 1.570796, 2.014841],accel_mss,speed_ms,0,blend_radius_m)
  movel([0.447686, -1.303085, -2.621295, -0.788010, 1.570796, 2.018482],accel_mss,speed_ms,0,blend_radius_m)
